--- program CFSteer (robot KUKA KR 30 HA) ---
  BAS (#INITMOV,0)
  BAS (#VEL_PTP,100)
  BAS (#ACC_PTP,20)
  Sollgeschwindigkeit (200.0 mm/s)
  Werkzeug setzen: TOOL 0
  Referenz erstellen.: BASE 0
  $ADVANCE = 5
  $APO.CPTP = 1.000
  $APO.CDIS = 1.000
  Sollgeschwindigkeit (1000.0 mm/s)
  Frame wechseln at (1415.36, -92.38, 659.99) mm, rotated rx -90 ry 0 rz 0 deg
  Werkzeug setzen at (350.64, -42.92, 173.8) mm
  Sollgeschwindigkeit (50.0 mm/s)
  MoveL 2 to (-32.85, -83.54, 62.24) mm, rotated rx 90 ry 17.84 rz 90 deg; joints [-6.49, -82.474, 137.961, 172.14, 55.739, -157.712]
  Sollgeschwindigkeit (50.0 mm/s)
  MoveL 3 to (-32.85, -40.71, 48.45) mm, rotated rx 90 ry 17.84 rz 90 deg; joints [-5.738, -79.848, 139.076, 173.33, 59.399, -158.749]
  MoveL 4 to (-31.86, -40.73, 48.38) mm, rotated rx 90 ry 17.46 rz 90 deg; joints [-5.612, -79.87, 138.999, 173.469, 59.293, -159.191]
  MoveL 5 to (-30.88, -40.75, 48.3) mm, rotated rx 90 ry 17.08 rz 90 deg; joints [-5.486, -79.891, 138.922, 173.609, 59.189, -159.635]
  MoveL 6 to (-29.89, -40.77, 48.23) mm, rotated rx 90 ry 16.7 rz 90 deg; joints [-5.359, -79.911, 138.845, 173.75, 59.085, -160.08]
  MoveL 7 to (-28.9, -40.8, 48.16) mm, rotated rx 90 ry 16.32 rz 90 deg; joints [-5.233, -79.929, 138.768, 173.891, 58.984, -160.524]
  MoveL 8 to (-27.92, -40.82, 48.09) mm, rotated rx 90 ry 15.94 rz 90 deg; joints [-5.106, -79.946, 138.691, 174.033, 58.883, -160.971]
  MoveL 9 to (-26.93, -40.84, 48.02) mm, rotated rx 90 ry 15.56 rz 90 deg; joints [-4.979, -79.961, 138.614, 174.175, 58.784, -161.417]
  MoveL 10 to (-25.95, -40.86, 47.95) mm, rotated rx 90 ry 15.17 rz 90 deg; joints [-4.852, -79.975, 138.537, 174.318, 58.687, -161.866]
  MoveL 11 to (-24.96, -40.88, 47.87) mm, rotated rx 90 ry 14.79 rz 90 deg; joints [-4.725, -79.988, 138.459, 174.461, 58.591, -162.314]
  MoveL 12 to (-23.97, -40.9, 47.8) mm, rotated rx 90 ry 14.41 rz 90 deg; joints [-4.598, -79.999, 138.382, 174.604, 58.496, -162.762]
  MoveL 13 to (-22.99, -40.9, 47.8) mm, rotated rx 90 ry 14.44 rz 90 deg; joints [-4.603, -79.938, 138.311, 174.598, 58.487, -162.729]
  MoveL 14 to (-22, -40.89, 47.81) mm, rotated rx 90 ry 14.47 rz 90 deg; joints [-4.608, -79.877, 138.24, 174.592, 58.478, -162.696]
  MoveL 15 to (-21.01, -40.89, 47.82) mm, rotated rx 90 ry 14.5 rz 90 deg; joints [-4.614, -79.815, 138.17, 174.585, 58.469, -162.663]
  MoveL 16 to (-20.02, -40.89, 47.82) mm, rotated rx 90 ry 14.53 rz 90 deg; joints [-4.618, -79.754, 138.099, 174.579, 58.459, -162.63]
  MoveL 17 to (-19.04, -40.89, 47.83) mm, rotated rx 90 ry 14.56 rz 90 deg; joints [-4.623, -79.693, 138.028, 174.572, 58.45, -162.597]
  MoveL 18 to (-18.05, -40.89, 47.83) mm, rotated rx 90 ry 14.59 rz 90 deg; joints [-4.628, -79.632, 137.957, 174.566, 58.44, -162.564]
  MoveL 19 to (-17.06, -40.89, 47.84) mm, rotated rx 90 ry 14.62 rz 90 deg; joints [-4.633, -79.571, 137.886, 174.56, 58.43, -162.53]
  MoveL 20 to (-16.07, -40.88, 47.84) mm, rotated rx 90 ry 14.64 rz 90 deg; joints [-4.638, -79.51, 137.815, 174.553, 58.421, -162.497]
  MoveL 21 to (-15.09, -40.88, 47.85) mm, rotated rx 90 ry 14.67 rz 90 deg; joints [-4.643, -79.449, 137.744, 174.547, 58.411, -162.464]
  MoveL 22 to (-14.11, -40.84, 47.99) mm, rotated rx 90 ry 15.42 rz 90 deg; joints [-4.875, -79.262, 137.685, 174.282, 58.551, -161.593]
  MoveL 23 to (-13.13, -40.8, 48.13) mm, rotated rx 90 ry 16.16 rz 90 deg; joints [-5.105, -79.07, 137.626, 174.022, 58.695, -160.725]
  MoveL 24 to (-12.15, -40.76, 48.27) mm, rotated rx 90 ry 16.9 rz 90 deg; joints [-5.334, -78.873, 137.566, 173.764, 58.843, -159.86]
  MoveL 25 to (-11.18, -40.72, 48.41) mm, rotated rx 90 ry 17.65 rz 90 deg; joints [-5.56, -78.673, 137.506, 173.509, 58.996, -158.998]
  MoveL 26 to (-10.2, -40.67, 48.55) mm, rotated rx 90 ry 18.39 rz 90 deg; joints [-5.785, -78.468, 137.446, 173.258, 59.153, -158.14]
  MoveL 27 to (-9.22, -40.63, 48.69) mm, rotated rx 90 ry 19.14 rz 90 deg; joints [-6.007, -78.259, 137.385, 173.01, 59.314, -157.285]
  MoveL 28 to (-8.24, -40.58, 48.83) mm, rotated rx 90 ry 19.88 rz 90 deg; joints [-6.228, -78.045, 137.323, 172.766, 59.479, -156.432]
  MoveL 29 to (-7.26, -40.53, 48.96) mm, rotated rx 90 ry 20.62 rz 90 deg; joints [-6.446, -77.828, 137.262, 172.525, 59.647, -155.585]
  MoveL 30 to (-6.28, -40.48, 49.1) mm, rotated rx 90 ry 21.37 rz 90 deg; joints [-6.662, -77.607, 137.2, 172.287, 59.82, -154.739]
  MoveL 31 to (-5.38, -40.38, 49.34) mm, rotated rx 90 ry 22.67 rz 90 deg; joints [-7.042, -77.252, 137.149, 171.874, 60.146, -153.264]
  MoveL 32 to (-4.47, -40.28, 49.57) mm, rotated rx 90 ry 23.98 rz 90 deg; joints [-7.415, -76.885, 137.096, 171.471, 60.485, -151.8]
  MoveL 33 to (-3.56, -40.17, 49.8) mm, rotated rx 90 ry 25.28 rz 90 deg; joints [-7.782, -76.505, 137.042, 171.079, 60.835, -150.347]
  MoveL 34 to (-2.66, -40.06, 50.03) mm, rotated rx 90 ry 26.58 rz 90 deg; joints [-8.143, -76.113, 136.987, 170.698, 61.196, -148.903]
  MoveL 35 to (-1.75, -39.94, 50.26) mm, rotated rx 90 ry 27.89 rz 90 deg; joints [-8.497, -75.708, 136.93, 170.327, 61.567, -147.472]
  MoveL 36 to (-0.84, -39.82, 50.49) mm, rotated rx 90 ry 29.19 rz 90 deg; joints [-8.844, -75.292, 136.872, 169.968, 61.948, -146.052]
  MoveL 37 to (0.05, -39.66, 50.77) mm, rotated rx 90 ry 30.83 rz 90 deg; joints [-9.272, -74.765, 136.814, 169.529, 62.446, -144.283]
  MoveL 38 to (0.93, -39.49, 51.04) mm, rotated rx 90 ry 32.47 rz 90 deg; joints [-9.689, -74.22, 136.754, 169.108, 62.958, -142.53]
  MoveL 39 to (1.82, -39.31, 51.31) mm, rotated rx 90 ry 34.11 rz 90 deg; joints [-10.094, -73.657, 136.691, 168.704, 63.484, -140.795]
  MoveL 40 to (2.71, -39.13, 51.57) mm, rotated rx 90 ry 35.75 rz 90 deg; joints [-10.488, -73.076, 136.624, 168.317, 64.023, -139.077]
  MoveL 41 to (3.6, -38.94, 51.83) mm, rotated rx 90 ry 37.39 rz 90 deg; joints [-10.87, -72.479, 136.554, 167.948, 64.574, -137.376]
  MoveL 42 to (4.49, -38.74, 52.08) mm, rotated rx 90 ry 39.02 rz 90 deg; joints [-11.239, -71.866, 136.481, 167.595, 65.136, -135.691]
  MoveL 43 to (5.36, -38.51, 52.36) mm, rotated rx 90 ry 40.85 rz 90 deg; joints [-11.636, -71.171, 136.404, 167.222, 65.775, -133.838]
  MoveL 44 to (6.24, -38.27, 52.62) mm, rotated rx 90 ry 42.67 rz 90 deg; joints [-12.018, -70.457, 136.322, 166.869, 66.426, -132.003]
  MoveL 45 to (7.12, -38.03, 52.88) mm, rotated rx 90 ry 44.49 rz 90 deg; joints [-12.383, -69.726, 136.235, 166.537, 67.088, -130.188]
  MoveL 46 to (7.99, -37.77, 53.13) mm, rotated rx 90 ry 46.31 rz 90 deg; joints [-12.733, -68.977, 136.144, 166.224, 67.759, -128.39]
  MoveL 47 to (8.87, -37.51, 53.38) mm, rotated rx 90 ry 48.13 rz 90 deg; joints [-13.066, -68.212, 136.047, 165.932, 68.438, -126.609]
  MoveL 48 to (9.75, -37.24, 53.61) mm, rotated rx 90 ry 49.95 rz 90 deg; joints [-13.383, -67.431, 135.945, 165.658, 69.125, -124.844]
  MoveL 49 to (10.62, -36.95, 53.85) mm, rotated rx 90 ry 51.84 rz 90 deg; joints [-13.694, -66.608, 135.837, 165.394, 69.846, -123.031]
  MoveL 50 to (11.5, -36.66, 54.07) mm, rotated rx 90 ry 53.73 rz 90 deg; joints [-13.987, -65.769, 135.723, 165.15, 70.572, -121.233]
  MoveL 51 to (12.37, -36.35, 54.28) mm, rotated rx 90 ry 55.62 rz 90 deg; joints [-14.261, -64.917, 135.603, 164.926, 71.303, -119.45]
  MoveL 52 to (13.24, -36.04, 54.49) mm, rotated rx 90 ry 57.5 rz 90 deg; joints [-14.518, -64.051, 135.476, 164.721, 72.039, -117.681]
  MoveL 53 to (14.12, -35.73, 54.68) mm, rotated rx 90 ry 59.39 rz 90 deg; joints [-14.755, -63.175, 135.344, 164.535, 72.776, -115.925]
  MoveL 54 to (14.99, -35.41, 54.87) mm, rotated rx 90 ry 61.28 rz 90 deg; joints [-14.974, -62.286, 135.206, 164.368, 73.517, -114.18]
  MoveL 55 to (15.87, -35.1, 55.03) mm, rotated rx 90 ry 63.05 rz 90 deg; joints [-15.161, -61.443, 135.067, 164.229, 74.209, -112.554]
  MoveL 56 to (16.74, -34.79, 55.18) mm, rotated rx 90 ry 64.82 rz 90 deg; joints [-15.332, -60.592, 134.922, 164.105, 74.901, -110.937]
  MoveL 57 to (17.61, -34.47, 55.32) mm, rotated rx 90 ry 66.59 rz 90 deg; joints [-15.486, -59.734, 134.772, 163.998, 75.593, -109.327]
  MoveL 58 to (18.49, -34.15, 55.46) mm, rotated rx 90 ry 68.36 rz 90 deg; joints [-15.624, -58.87, 134.616, 163.905, 76.283, -107.725]
  MoveL 59 to (19.36, -33.82, 55.58) mm, rotated rx 90 ry 70.13 rz 90 deg; joints [-15.744, -58.001, 134.456, 163.829, 76.972, -106.129]
  MoveL 60 to (20.23, -33.49, 55.69) mm, rotated rx 90 ry 71.9 rz 90 deg; joints [-15.848, -57.128, 134.289, 163.767, 77.657, -104.538]
  MoveL 61 to (21.12, -33.23, 55.78) mm, rotated rx 90 ry 73.31 rz 90 deg; joints [-15.916, -56.424, 134.139, 163.73, 78.193, -103.273]
  MoveL 62 to (22, -32.97, 55.85) mm, rotated rx 90 ry 74.72 rz 90 deg; joints [-15.973, -55.719, 133.986, 163.704, 78.726, -102.01]
  MoveL 63 to (22.88, -32.7, 55.92) mm, rotated rx 90 ry 76.13 rz 90 deg; joints [-16.02, -55.013, 133.83, 163.686, 79.256, -100.749]
  MoveL 64 to (23.77, -32.43, 55.98) mm, rotated rx 90 ry 77.54 rz 90 deg; joints [-16.056, -54.307, 133.67, 163.678, 79.783, -99.49]
  MoveL 65 to (24.65, -32.16, 56.04) mm, rotated rx 90 ry 78.95 rz 90 deg; joints [-16.082, -53.6, 133.508, 163.679, 80.307, -98.231]
  MoveL 66 to (25.53, -31.89, 56.09) mm, rotated rx 90 ry 80.36 rz 90 deg; joints [-16.096, -52.893, 133.342, 163.689, 80.827, -96.974]
  MoveL 67 to (26.46, -31.75, 56.11) mm, rotated rx 90 ry 81.07 rz 90 deg; joints [-16.093, -52.524, 133.222, 163.704, 81.065, -96.333]
  MoveL 68 to (27.39, -31.61, 56.13) mm, rotated rx 90 ry 81.78 rz 90 deg; joints [-16.087, -52.155, 133.1, 163.721, 81.303, -95.692]
  MoveL 69 to (28.32, -31.47, 56.15) mm, rotated rx 90 ry 82.49 rz 90 deg; joints [-16.078, -51.786, 132.978, 163.74, 81.539, -95.051]
  MoveL 70 to (29.25, -31.33, 56.17) mm, rotated rx 90 ry 83.2 rz 90 deg; joints [-16.067, -51.418, 132.856, 163.762, 81.774, -94.409]
  MoveL 71 to (30.18, -31.19, 56.19) mm, rotated rx 90 ry 83.92 rz 90 deg; joints [-16.053, -51.052, 132.733, 163.785, 82.008, -93.768]
  MoveL 72 to (31.11, -31.05, 56.2) mm, rotated rx 90 ry 84.63 rz 90 deg; joints [-16.036, -50.685, 132.608, 163.812, 82.24, -93.125]
  MoveL 73 to (31.98, -31.11, 56.2) mm, rotated rx 90 ry 84.31 rz 90 deg; joints [-16.026, -50.818, 132.569, 163.815, 82.074, -93.398]
  MoveL 74 to (32.86, -31.18, 56.19) mm, rotated rx 90 ry 83.99 rz 90 deg; joints [-16.016, -50.951, 132.53, 163.819, 81.907, -93.671]
  MoveL 75 to (33.73, -31.24, 56.18) mm, rotated rx 90 ry 83.67 rz 90 deg; joints [-16.005, -51.084, 132.49, 163.823, 81.742, -93.943]
  MoveL 76 to (34.6, -31.3, 56.17) mm, rotated rx 90 ry 83.35 rz 90 deg; joints [-15.993, -51.216, 132.45, 163.828, 81.576, -94.216]
  MoveL 77 to (35.48, -31.36, 56.17) mm, rotated rx 90 ry 83.03 rz 90 deg; joints [-15.981, -51.348, 132.41, 163.833, 81.41, -94.489]
  MoveL 78 to (36.35, -31.43, 56.16) mm, rotated rx 90 ry 82.71 rz 90 deg; joints [-15.968, -51.479, 132.37, 163.838, 81.245, -94.762]
  MoveL 79 to (37.22, -31.49, 56.15) mm, rotated rx 90 ry 82.39 rz 90 deg; joints [-15.955, -51.61, 132.329, 163.844, 81.079, -95.035]
  MoveL 80 to (38.14, -31.69, 56.12) mm, rotated rx 90 ry 81.34 rz 90 deg; joints [-15.935, -52.089, 132.339, 163.843, 80.628, -95.954]
  MoveL 81 to (39.06, -31.9, 56.09) mm, rotated rx 90 ry 80.3 rz 90 deg; joints [-15.909, -52.566, 132.346, 163.847, 80.176, -96.874]
  MoveL 82 to (39.98, -32.1, 56.05) mm, rotated rx 90 ry 79.25 rz 90 deg; joints [-15.878, -53.042, 132.353, 163.856, 79.723, -97.796]
  MoveL 83 to (40.9, -32.3, 56.01) mm, rotated rx 90 ry 78.2 rz 90 deg; joints [-15.84, -53.516, 132.357, 163.87, 79.27, -98.718]
  MoveL 84 to (41.81, -32.5, 55.97) mm, rotated rx 90 ry 77.15 rz 90 deg; joints [-15.797, -53.988, 132.359, 163.889, 78.816, -99.641]
  MoveL 85 to (42.73, -32.7, 55.92) mm, rotated rx 90 ry 76.1 rz 90 deg; joints [-15.748, -54.458, 132.36, 163.912, 78.362, -100.566]
  MoveL 86 to (43.65, -32.9, 55.87) mm, rotated rx 90 ry 75.06 rz 90 deg; joints [-15.694, -54.926, 132.358, 163.941, 77.908, -101.493]
  MoveL 87 to (44.61, -32.99, 55.84) mm, rotated rx 90 ry 74.56 rz 90 deg; joints [-15.659, -55.131, 132.318, 163.962, 77.67, -101.928]
  MoveL 88 to (45.57, -33.09, 55.82) mm, rotated rx 90 ry 74.06 rz 90 deg; joints [-15.623, -55.336, 132.277, 163.984, 77.432, -102.364]
  MoveL 89 to (46.52, -33.18, 55.79) mm, rotated rx 90 ry 73.56 rz 90 deg; joints [-15.585, -55.54, 132.236, 164.007, 77.194, -102.8]
  MoveL 90 to (47.48, -33.28, 55.76) mm, rotated rx 90 ry 73.07 rz 90 deg; joints [-15.547, -55.742, 132.194, 164.031, 76.956, -103.236]
  MoveL 91 to (48.44, -33.37, 55.73) mm, rotated rx 90 ry 72.57 rz 90 deg; joints [-15.507, -55.944, 132.152, 164.056, 76.719, -103.673]
  MoveL 92 to (49.4, -33.46, 55.7) mm, rotated rx 90 ry 72.08 rz 90 deg; joints [-15.466, -56.145, 132.109, 164.082, 76.482, -104.111]
  MoveL 93 to (50.35, -33.55, 55.67) mm, rotated rx 90 ry 71.58 rz 90 deg; joints [-15.424, -56.345, 132.066, 164.109, 76.245, -104.55]
  MoveL 94 to (51.31, -33.44, 55.71) mm, rotated rx 90 ry 72.18 rz 90 deg; joints [-15.447, -56.037, 131.96, 164.099, 76.442, -103.999]
  MoveL 95 to (52.26, -33.33, 55.75) mm, rotated rx 90 ry 72.78 rz 90 deg; joints [-15.468, -55.728, 131.853, 164.09, 76.638, -103.448]
  MoveL 96 to (53.21, -33.22, 55.78) mm, rotated rx 90 ry 73.39 rz 90 deg; joints [-15.488, -55.419, 131.746, 164.083, 76.832, -102.898]
  MoveL 97 to (54.16, -33.1, 55.81) mm, rotated rx 90 ry 73.99 rz 90 deg; joints [-15.505, -55.11, 131.638, 164.078, 77.027, -102.348]
  MoveL 98 to (55.12, -32.99, 55.85) mm, rotated rx 90 ry 74.59 rz 90 deg; joints [-15.521, -54.802, 131.53, 164.074, 77.221, -101.798]
  MoveL 99 to (56.07, -32.88, 55.88) mm, rotated rx 90 ry 75.19 rz 90 deg; joints [-15.535, -54.493, 131.421, 164.073, 77.414, -101.249]
  MoveL 100 to (57.02, -32.76, 55.91) mm, rotated rx 90 ry 75.8 rz 90 deg; joints [-15.547, -54.185, 131.312, 164.073, 77.605, -100.7]
  MoveL 101 to (57.94, -32.56, 55.95) mm, rotated rx 90 ry 76.82 rz 90 deg; joints [-15.572, -53.681, 131.177, 164.069, 77.962, -99.772]
  MoveL 102 to (58.86, -32.37, 56) mm, rotated rx 90 ry 77.85 rz 90 deg; joints [-15.591, -53.177, 131.04, 164.07, 78.317, -98.846]
  MoveL 103 to (59.77, -32.17, 56.04) mm, rotated rx 90 ry 78.87 rz 90 deg; joints [-15.605, -52.672, 130.902, 164.076, 78.67, -97.92]
  MoveL 104 to (60.69, -31.97, 56.08) mm, rotated rx 90 ry 79.9 rz 90 deg; joints [-15.614, -52.169, 130.763, 164.087, 79.02, -96.995]
  MoveL 105 to (61.61, -31.77, 56.11) mm, rotated rx 90 ry 80.92 rz 90 deg; joints [-15.617, -51.665, 130.622, 164.103, 79.369, -96.069]
  MoveL 106 to (62.52, -31.58, 56.14) mm, rotated rx 90 ry 81.95 rz 90 deg; joints [-15.614, -51.163, 130.48, 164.124, 79.715, -95.145]
  MoveL 107 to (63.44, -31.38, 56.17) mm, rotated rx 90 ry 82.97 rz 90 deg; joints [-15.607, -50.661, 130.336, 164.149, 80.06, -94.22]
  MoveL 108 to (64.31, -31.34, 56.17) mm, rotated rx 90 ry 83.18 rz 90 deg; joints [-15.596, -50.54, 130.255, 164.162, 80.098, -94.022]
  MoveL 109 to (65.17, -31.29, 56.17) mm, rotated rx 90 ry 83.4 rz 90 deg; joints [-15.584, -50.42, 130.175, 164.176, 80.136, -93.825]
  MoveL 110 to (66.03, -31.25, 56.18) mm, rotated rx 90 ry 83.61 rz 90 deg; joints [-15.573, -50.299, 130.094, 164.19, 80.174, -93.627]
  MoveL 111 to (66.9, -31.21, 56.19) mm, rotated rx 90 ry 83.82 rz 90 deg; joints [-15.561, -50.179, 130.014, 164.203, 80.211, -93.429]
  MoveL 112 to (67.76, -31.17, 56.19) mm, rotated rx 90 ry 84.03 rz 90 deg; joints [-15.549, -50.058, 129.933, 164.217, 80.249, -93.231]
  MoveL 113 to (68.63, -31.13, 56.19) mm, rotated rx 90 ry 84.24 rz 90 deg; joints [-15.537, -49.938, 129.853, 164.232, 80.286, -93.033]
  MoveL 114 to (69.49, -31.09, 56.2) mm, rotated rx 90 ry 84.45 rz 90 deg; joints [-15.524, -49.819, 129.772, 164.246, 80.323, -92.835]
  MoveL 115 to (70.41, -31.25, 56.18) mm, rotated rx 90 ry 83.65 rz 90 deg; joints [-15.516, -50.166, 129.763, 164.238, 79.98, -93.541]
  MoveL 116 to (71.33, -31.4, 56.16) mm, rotated rx 90 ry 82.84 rz 90 deg; joints [-15.504, -50.513, 129.753, 164.232, 79.637, -94.248]
  MoveL 117 to (72.26, -31.56, 56.14) mm, rotated rx 90 ry 82.04 rz 90 deg; joints [-15.489, -50.859, 129.743, 164.23, 79.292, -94.955]
  MoveL 118 to (73.18, -31.71, 56.12) mm, rotated rx 90 ry 81.24 rz 90 deg; joints [-15.47, -51.204, 129.731, 164.23, 78.948, -95.664]
  MoveL 119 to (74.1, -31.87, 56.09) mm, rotated rx 90 ry 80.43 rz 90 deg; joints [-15.448, -51.549, 129.718, 164.233, 78.603, -96.373]
  MoveL 120 to (75.03, -32.02, 56.07) mm, rotated rx 90 ry 79.63 rz 90 deg; joints [-15.423, -51.892, 129.704, 164.239, 78.258, -97.082]
  MoveL 121 to (75.91, -32.31, 56.01) mm, rotated rx 90 ry 78.17 rz 90 deg; joints [-15.379, -52.536, 129.737, 164.248, 77.667, -98.381]
  MoveL 122 to (76.79, -32.59, 55.95) mm, rotated rx 90 ry 76.71 rz 90 deg; joints [-15.325, -53.177, 129.765, 164.267, 77.074, -99.683]
  MoveL 123 to (77.67, -32.86, 55.88) mm, rotated rx 90 ry 75.25 rz 90 deg; joints [-15.259, -53.814, 129.791, 164.295, 76.48, -100.988]
  MoveL 124 to (78.55, -33.14, 55.8) mm, rotated rx 90 ry 73.79 rz 90 deg; joints [-15.183, -54.449, 129.813, 164.333, 75.886, -102.297]
  MoveL 125 to (79.43, -33.41, 55.72) mm, rotated rx 90 ry 72.33 rz 90 deg; joints [-15.095, -55.079, 129.831, 164.38, 75.291, -103.61]
  MoveL 126 to (80.31, -33.69, 55.63) mm, rotated rx 90 ry 70.87 rz 90 deg; joints [-14.997, -55.704, 129.846, 164.438, 74.696, -104.926]
  MoveL 127 to (81.19, -34.02, 55.51) mm, rotated rx 90 ry 69.08 rz 90 deg; joints [-14.865, -56.471, 129.876, 164.519, 73.975, -106.551]
  MoveL 128 to (82.06, -34.34, 55.38) mm, rotated rx 90 ry 67.28 rz 90 deg; joints [-14.717, -57.231, 129.9, 164.616, 73.255, -108.183]
  MoveL 129 to (82.93, -34.67, 55.24) mm, rotated rx 90 ry 65.49 rz 90 deg; joints [-14.553, -57.982, 129.919, 164.727, 72.536, -109.824]
  MoveL 130 to (83.81, -34.98, 55.09) mm, rotated rx 90 ry 63.7 rz 90 deg; joints [-14.373, -58.723, 129.933, 164.855, 71.819, -111.475]
  MoveL 131 to (84.68, -35.3, 54.92) mm, rotated rx 90 ry 61.91 rz 90 deg; joints [-14.177, -59.453, 129.941, 164.997, 71.105, -113.135]
  MoveL 132 to (85.55, -35.61, 54.75) mm, rotated rx 90 ry 60.11 rz 90 deg; joints [-13.966, -60.173, 129.945, 165.156, 70.394, -114.807]
  MoveL 133 to (86.51, -35.95, 54.55) mm, rotated rx 90 ry 58.07 rz 90 deg; joints [-13.706, -60.981, 129.945, 165.356, 69.59, -116.727]
  MoveL 134 to (87.46, -36.29, 54.33) mm, rotated rx 90 ry 56.02 rz 90 deg; joints [-13.427, -61.772, 129.939, 165.577, 68.793, -118.664]
  MoveL 135 to (88.42, -36.62, 54.1) mm, rotated rx 90 ry 53.98 rz 90 deg; joints [-13.129, -62.546, 129.926, 165.82, 68.003, -120.618]
  MoveL 136 to (89.37, -36.94, 53.86) mm, rotated rx 90 ry 51.93 rz 90 deg; joints [-12.811, -63.301, 129.907, 166.085, 67.222, -122.59]
  MoveL 137 to (90.32, -37.25, 53.6) mm, rotated rx 90 ry 49.89 rz 90 deg; joints [-12.474, -64.036, 129.882, 166.372, 66.451, -124.581]
  MoveL 138 to (91.28, -37.55, 53.34) mm, rotated rx 90 ry 47.84 rz 90 deg; joints [-12.119, -64.751, 129.851, 166.682, 65.691, -126.593]
  MoveL 139 to (92.23, -37.84, 53.06) mm, rotated rx 90 ry 45.8 rz 90 deg; joints [-11.745, -65.445, 129.814, 167.014, 64.943, -128.626]
  MoveL 140 to (93.19, -38.13, 52.78) mm, rotated rx 90 ry 43.75 rz 90 deg; joints [-11.354, -66.116, 129.771, 167.37, 64.209, -130.681]
  MoveL 141 to (94.15, -38.37, 52.52) mm, rotated rx 90 ry 41.92 rz 90 deg; joints [-10.987, -66.693, 129.719, 167.711, 63.559, -132.544]
  MoveL 142 to (95.12, -38.61, 52.24) mm, rotated rx 90 ry 40.08 rz 90 deg; joints [-10.606, -67.25, 129.663, 168.07, 62.923, -134.426]
  MoveL 143 to (96.08, -38.84, 51.96) mm, rotated rx 90 ry 38.25 rz 90 deg; joints [-10.212, -67.788, 129.603, 168.449, 62.3, -136.327]
  MoveL 144 to (97.05, -39.05, 51.68) mm, rotated rx 90 ry 36.41 rz 90 deg; joints [-9.805, -68.305, 129.539, 168.847, 61.693, -138.248]
  MoveL 145 to (98.01, -39.26, 51.38) mm, rotated rx 90 ry 34.58 rz 90 deg; joints [-9.386, -68.8, 129.471, 169.264, 61.102, -140.188]
  MoveL 146 to (98.98, -39.46, 51.09) mm, rotated rx 90 ry 32.74 rz 90 deg; joints [-8.955, -69.274, 129.4, 169.7, 60.527, -142.149]
  MoveL 147 to (99.94, -39.65, 50.78) mm, rotated rx 90 ry 30.91 rz 90 deg; joints [-8.512, -69.725, 129.326, 170.156, 59.97, -144.13]
  MoveL 148 to (100.91, -39.83, 50.47) mm, rotated rx 90 ry 29.07 rz 90 deg; joints [-8.057, -70.154, 129.248, 170.631, 59.431, -146.132]
  MoveL 149 to (101.91, -39.95, 50.24) mm, rotated rx 90 ry 27.77 rz 90 deg; joints [-7.727, -70.429, 129.167, 170.981, 59.053, -147.563]
  MoveL 150 to (102.9, -40.07, 50.01) mm, rotated rx 90 ry 26.47 rz 90 deg; joints [-7.391, -70.691, 129.085, 171.34, 58.686, -149.004]
  MoveL 151 to (103.9, -40.18, 49.78) mm, rotated rx 90 ry 25.17 rz 90 deg; joints [-7.05, -70.942, 129.001, 171.709, 58.329, -150.457]
  MoveL 152 to (104.89, -40.29, 49.55) mm, rotated rx 90 ry 23.87 rz 90 deg; joints [-6.704, -71.18, 128.916, 172.086, 57.983, -151.918]
  MoveL 153 to (105.89, -40.39, 49.32) mm, rotated rx 90 ry 22.57 rz 90 deg; joints [-6.354, -71.406, 128.829, 172.472, 57.649, -153.389]
  MoveL 154 to (106.89, -40.48, 49.08) mm, rotated rx 90 ry 21.26 rz 90 deg; joints [-6, -71.619, 128.742, 172.866, 57.326, -154.87]
  MoveL 155 to (107.88, -40.57, 48.84) mm, rotated rx 90 ry 19.96 rz 90 deg; joints [-5.642, -71.82, 128.653, 173.269, 57.015, -156.36]
  MoveL 156 to (108.88, -40.66, 48.6) mm, rotated rx 90 ry 18.66 rz 90 deg; joints [-5.28, -72.008, 128.564, 173.68, 56.716, -157.859]
  MoveL 157 to (109.79, -40.69, 48.51) mm, rotated rx 90 ry 18.16 rz 90 deg; joints [-5.135, -72.05, 128.488, 173.845, 56.591, -158.446]
  MoveL 158 to (110.7, -40.72, 48.41) mm, rotated rx 90 ry 17.65 rz 90 deg; joints [-4.99, -72.091, 128.413, 174.01, 56.467, -159.035]
  MoveL 159 to (111.61, -40.75, 48.32) mm, rotated rx 90 ry 17.14 rz 90 deg; joints [-4.845, -72.129, 128.337, 174.176, 56.345, -159.624]
  MoveL 160 to (112.52, -40.78, 48.22) mm, rotated rx 90 ry 16.63 rz 90 deg; joints [-4.699, -72.165, 128.262, 174.344, 56.226, -160.215]
  MoveL 161 to (113.43, -40.81, 48.12) mm, rotated rx 90 ry 16.13 rz 90 deg; joints [-4.553, -72.199, 128.186, 174.512, 56.108, -160.806]
  MoveL 162 to (114.34, -40.84, 48.03) mm, rotated rx 90 ry 15.62 rz 90 deg; joints [-4.407, -72.232, 128.11, 174.682, 55.992, -161.401]
  MoveL 163 to (115.25, -40.86, 47.93) mm, rotated rx 90 ry 15.11 rz 90 deg; joints [-4.26, -72.262, 128.033, 174.852, 55.879, -161.995]
  MoveL 164 to (116.16, -40.89, 47.84) mm, rotated rx 90 ry 14.61 rz 90 deg; joints [-4.113, -72.29, 127.957, 175.024, 55.768, -162.591]
  MoveL 165 to (117.07, -40.91, 47.74) mm, rotated rx 90 ry 14.1 rz 90 deg; joints [-3.965, -72.316, 127.88, 175.196, 55.658, -163.187]
  MoveL 166 to (117.99, -40.91, 47.76) mm, rotated rx 90 ry 14.17 rz 90 deg; joints [-3.984, -72.256, 127.811, 175.172, 55.65, -163.097]
  MoveL 167 to (118.9, -40.9, 47.77) mm, rotated rx 90 ry 14.25 rz 90 deg; joints [-4.003, -72.197, 127.742, 175.149, 55.641, -163.006]
  MoveL 168 to (119.81, -40.9, 47.78) mm, rotated rx 90 ry 14.33 rz 90 deg; joints [-4.022, -72.137, 127.673, 175.126, 55.633, -162.915]
  MoveL 169 to (120.73, -40.9, 47.8) mm, rotated rx 90 ry 14.41 rz 90 deg; joints [-4.041, -72.077, 127.603, 175.102, 55.624, -162.824]
  MoveL 170 to (121.64, -40.89, 47.81) mm, rotated rx 90 ry 14.48 rz 90 deg; joints [-4.059, -72.017, 127.534, 175.079, 55.616, -162.733]
  MoveL 171 to (122.55, -40.89, 47.83) mm, rotated rx 90 ry 14.56 rz 90 deg; joints [-4.078, -71.957, 127.464, 175.056, 55.607, -162.643]
  MoveL 172 to (123.47, -40.88, 47.84) mm, rotated rx 90 ry 14.64 rz 90 deg; joints [-4.097, -71.897, 127.395, 175.033, 55.598, -162.552]
  MoveL 173 to (124.38, -40.88, 47.86) mm, rotated rx 90 ry 14.71 rz 90 deg; joints [-4.116, -71.837, 127.326, 175.009, 55.59, -162.46]
  MoveL 174 to (125.3, -40.88, 47.87) mm, rotated rx 90 ry 14.79 rz 90 deg; joints [-4.134, -71.777, 127.256, 174.986, 55.581, -162.369]
  MoveL 175 to (126.21, -40.86, 47.94) mm, rotated rx 90 ry 15.16 rz 90 deg; joints [-4.235, -71.673, 127.19, 174.867, 55.624, -161.934]
  MoveL 176 to (127.12, -40.84, 48.01) mm, rotated rx 90 ry 15.53 rz 90 deg; joints [-4.336, -71.568, 127.124, 174.747, 55.668, -161.499]
  MoveL 177 to (128.03, -40.82, 48.08) mm, rotated rx 90 ry 15.9 rz 90 deg; joints [-4.436, -71.462, 127.058, 174.629, 55.713, -161.064]
  MoveL 178 to (128.94, -40.8, 48.15) mm, rotated rx 90 ry 16.27 rz 90 deg; joints [-4.536, -71.356, 126.992, 174.511, 55.759, -160.63]
  MoveL 179 to (129.86, -40.78, 48.22) mm, rotated rx 90 ry 16.64 rz 90 deg; joints [-4.635, -71.248, 126.926, 174.394, 55.805, -160.197]
  MoveL 180 to (130.77, -40.76, 48.29) mm, rotated rx 90 ry 17.02 rz 90 deg; joints [-4.734, -71.14, 126.859, 174.277, 55.852, -159.764]
  MoveL 181 to (131.68, -40.74, 48.36) mm, rotated rx 90 ry 17.39 rz 90 deg; joints [-4.832, -71.031, 126.793, 174.161, 55.9, -159.332]
  MoveL 182 to (132.59, -40.71, 48.43) mm, rotated rx 90 ry 17.76 rz 90 deg; joints [-4.93, -70.921, 126.726, 174.046, 55.949, -158.9]
  MoveL 183 to (133.51, -40.69, 48.5) mm, rotated rx 90 ry 18.13 rz 90 deg; joints [-5.027, -70.81, 126.659, 173.932, 55.999, -158.469]
  MoveL 184 to (134.42, -40.67, 48.56) mm, rotated rx 90 ry 18.43 rz 90 deg; joints [-5.106, -70.71, 126.591, 173.84, 56.035, -158.119]
  MoveL 185 to (135.33, -40.65, 48.61) mm, rotated rx 90 ry 18.73 rz 90 deg; joints [-5.184, -70.609, 126.524, 173.749, 56.073, -157.767]
  MoveL 186 to (136.25, -40.63, 48.67) mm, rotated rx 90 ry 19.04 rz 90 deg; joints [-5.262, -70.508, 126.456, 173.657, 56.11, -157.416]
  MoveL 187 to (137.16, -40.62, 48.73) mm, rotated rx 90 ry 19.34 rz 90 deg; joints [-5.339, -70.407, 126.388, 173.567, 56.149, -157.066]
  MoveL 188 to (138.07, -40.59, 48.78) mm, rotated rx 90 ry 19.64 rz 90 deg; joints [-5.416, -70.305, 126.32, 173.477, 56.187, -156.716]
  MoveL 189 to (138.98, -40.58, 48.84) mm, rotated rx 90 ry 19.95 rz 90 deg; joints [-5.493, -70.202, 126.252, 173.387, 56.226, -156.366]
  MoveL 190 to (139.9, -40.55, 48.89) mm, rotated rx 90 ry 20.25 rz 90 deg; joints [-5.57, -70.099, 126.183, 173.298, 56.266, -156.017]
  MoveL 191 to (140.81, -40.53, 48.95) mm, rotated rx 90 ry 20.55 rz 90 deg; joints [-5.646, -69.996, 126.115, 173.21, 56.306, -155.669]
  MoveL 192 to (141.72, -40.51, 49.01) mm, rotated rx 90 ry 20.85 rz 90 deg; joints [-5.721, -69.892, 126.047, 173.122, 56.346, -155.322]
  MoveL 193 to (142.4, -40.79, 48.17) mm, rotated rx 90 ry 16.38 rz 90 deg; joints [-4.515, -70.63, 125.949, 174.515, 55.442, -160.499]
  MoveL 194 to (143.07, -41.01, 47.32) mm, rotated rx 90 ry 11.91 rz 90 deg; joints [-3.266, -71.227, 125.841, 175.996, 54.68, -165.771]
  MoveL 195 to (143.75, -41.16, 46.46) mm, rotated rx 90 ry 7.44 rz 90 deg; joints [-1.981, -71.678, 125.723, 177.553, 54.07, -171.124]
  MoveL 196 to (144.43, -41.23, 45.58) mm, rotated rx 90 ry 2.97 rz 90 deg; joints [-0.67, -71.982, 125.598, 179.168, 53.619, -176.537]
  MoveL 197 to (145.1, -41.25, 44.7) mm, rotated rx 90 ry 0 rz 90 deg; joints [0.224, -72.088, 125.494, -179.721, 53.406, 179.834]
  MoveL 198 to (141.7, -41.25, 42.87) mm, rotated rx 90 ry 0 rz 90 deg; joints [0.311, -72.273, 125.758, -179.612, 53.486, 179.769]
  MoveL 199 to (137.91, -41.25, 41.96) mm, rotated rx 90 ry 0 rz 90 deg; joints [0.355, -72.478, 126.051, -179.558, 53.573, 179.738]
  MoveL 200 to (134, -41.25, 41.48) mm, rotated rx 90 ry 0 rz 90 deg; joints [0.379, -72.691, 126.353, -179.529, 53.663, 179.721]
  MoveL 201 to (130.09, -41.25, 41.08) mm, rotated rx 90 ry 0 rz 90 deg; joints [0.4, -72.903, 126.655, -179.505, 53.752, 179.707]
  MoveL 202 to (126.21, -41.25, 40.71) mm, rotated rx 90 ry 0 rz 90 deg; joints [0.419, -73.115, 126.954, -179.481, 53.84, 179.694]
  MoveL 203 to (118.64, -41.25, 39.88) mm, rotated rx 90 ry 0 rz 90 deg; joints [0.461, -73.528, 127.535, -179.43, 54.008, 179.665]
  MoveL 204 to (111.13, -41.25, 38.67) mm, rotated rx 90 ry 0 rz 90 deg; joints [0.523, -73.939, 128.109, -179.355, 54.172, 179.623]
  MoveL 205 to (104.5, -41.25, 37.04) mm, rotated rx 90 ry 0 rz 90 deg; joints [0.605, -74.302, 128.613, -179.255, 54.314, 179.565]
  MoveL 206 to (98.04, -41.25, 34.74) mm, rotated rx 90 ry 0 rz 90 deg; joints [0.721, -74.656, 129.102, -179.113, 54.45, 179.485]
  MoveL 207 to (91.88, -41.25, 31.62) mm, rotated rx 90 ry 0 rz 90 deg; joints [0.879, -74.993, 129.566, -178.922, 54.578, 179.375]
  MoveL 208 to (86.28, -41.25, 27.66) mm, rotated rx 90 ry 0 rz 90 deg; joints [1.079, -75.299, 129.984, -178.678, 54.692, 179.236]
  MoveL 209 to (80.96, -41.25, 22.17) mm, rotated rx 90 ry 0 rz 90 deg; joints [1.356, -75.587, 130.376, -178.34, 54.801, 179.043]
  MoveL 210 to (76.3, -41.25, 15.86) mm, rotated rx 90 ry 0 rz 90 deg; joints [1.677, -75.837, 130.714, -177.95, 54.895, 178.821]
  MoveL 211 to (75.7, -41.25, 15.02) mm, rotated rx 90 ry 0 rz 90 deg; joints [1.72, -75.868, 130.757, -177.898, 54.907, 178.791]
  MoveL 212 to (75.11, -41.22, 14.18) mm, rotated rx 90 ry -4.2 rz 90 deg; joints [3.049, -75.959, 130.67, -176.267, 54.768, 173.646]
  MoveL 213 to (74.51, -41.13, 13.34) mm, rotated rx 90 ry -8.49 rz 90 deg; joints [4.409, -75.905, 130.577, -174.602, 54.792, 168.391]
  MoveL 214 to (73.92, -40.97, 12.51) mm, rotated rx 90 ry -12.78 rz 90 deg; joints [5.762, -75.702, 130.481, -172.958, 54.983, 163.164]
  MoveL 215 to (73.33, -40.76, 11.71) mm, rotated rx 90 ry -17.03 rz 90 deg; joints [7.085, -75.358, 130.384, -171.375, 55.332, 158.042]
  MoveL 216 to (72.75, -40.48, 10.92) mm, rotated rx 90 ry -21.27 rz 90 deg; joints [8.385, -74.874, 130.285, -169.849, 55.833, 152.988]
  MoveL 217 to (72.17, -40.15, 10.15) mm, rotated rx 90 ry -25.52 rz 90 deg; joints [9.653, -74.253, 130.184, -168.397, 56.477, 148.015]
  MoveL 218 to (71.58, -39.77, 9.42) mm, rotated rx 90 ry -29.76 rz 90 deg; joints [10.881, -73.501, 130.08, -167.03, 57.256, 143.14]
  MoveL 219 to (71.04, -39.35, 8.74) mm, rotated rx 90 ry -33.79 rz 90 deg; joints [12.006, -72.668, 129.976, -165.819, 58.109, 138.604]
  MoveL 220 to (70.5, -38.89, 8.1) mm, rotated rx 90 ry -37.83 rz 90 deg; joints [13.083, -71.724, 129.868, -164.698, 59.064, 134.168]
  MoveL 221 to (69.96, -38.38, 7.49) mm, rotated rx 90 ry -41.86 rz 90 deg; joints [14.108, -70.676, 129.755, -163.671, 60.109, 129.834]
  MoveL 222 to (69.42, -37.83, 6.92) mm, rotated rx 90 ry -45.89 rz 90 deg; joints [15.077, -69.53, 129.636, -162.739, 61.234, 125.604]
  MoveL 223 to (68.95, -37.22, 6.38) mm, rotated rx 90 ry -50.05 rz 90 deg; joints [16.009, -68.247, 129.499, -161.879, 62.464, 121.349]
  MoveL 224 to (68.49, -36.58, 5.88) mm, rotated rx 90 ry -54.2 rz 90 deg; joints [16.874, -66.873, 129.353, -161.118, 63.758, 117.196]
  MoveL 225 to (68.02, -35.9, 5.42) mm, rotated rx 90 ry -58.36 rz 90 deg; joints [17.667, -65.415, 129.197, -160.453, 65.105, 113.14]
  MoveL 226 to (67.55, -35.19, 5.02) mm, rotated rx 90 ry -62.52 rz 90 deg; joints [18.386, -63.882, 129.03, -159.882, 66.495, 109.172]
  MoveL 227 to (67.13, -34.29, 4.6) mm, rotated rx 90 ry -67.57 rz 90 deg; joints [19.155, -61.92, 128.8, -159.309, 68.228, 104.454]
  MoveL 228 to (66.72, -33.36, 4.26) mm, rotated rx 90 ry -72.63 rz 90 deg; joints [19.807, -59.872, 128.552, -158.863, 69.997, 99.839]
  MoveL 229 to (66.3, -32.4, 4.01) mm, rotated rx 90 ry -77.68 rz 90 deg; joints [20.339, -57.755, 128.286, -158.537, 71.79, 95.311]
  MoveL 230 to (65.88, -31.42, 3.84) mm, rotated rx 90 ry -82.74 rz 90 deg; joints [20.751, -55.583, 128.002, -158.325, 73.593, 90.855]
  MoveL 231 to (65.46, -30.43, 3.76) mm, rotated rx 90 ry -87.8 rz 90 deg; joints [21.039, -53.372, 127.701, -158.223, 75.397, 86.453]
  MoveL 232 to (65.15, -29.59, 3.75) mm, rotated rx 0 ry -90 rz 180 deg; joints [21.129, -52.375, 127.571, -158.213, 76.211, 84.558]
  MoveL 233 to (64.83, -28.74, 3.75) mm, rotated rx 0 ry -90 rz 180 deg; joints [21.134, -52.326, 127.587, -158.213, 76.273, 84.582]
  MoveL 234 to (64.52, -27.89, 3.75) mm, rotated rx 0 ry -90 rz 180 deg; joints [21.139, -52.277, 127.604, -158.214, 76.334, 84.606]
  MoveL 235 to (64.21, -27.04, 3.75) mm, rotated rx 0 ry -90 rz 180 deg; joints [21.145, -52.227, 127.62, -158.214, 76.396, 84.629]
  MoveL 236 to (63.9, -26.19, 3.75) mm, rotated rx 0 ry -90 rz 180 deg; joints [21.15, -52.178, 127.637, -158.215, 76.458, 84.653]
  MoveL 237 to (63.59, -25.34, 3.75) mm, rotated rx 0 ry -90 rz 180 deg; joints [21.155, -52.128, 127.653, -158.215, 76.519, 84.677]
  MoveL 238 to (61.65, -20.55, 3.75) mm, rotated rx 0 ry -90 rz 180 deg; joints [21.188, -51.853, 127.757, -158.215, 76.875, 84.814]
  MoveL 239 to (59.77, -17.22, 3.75) mm, rotated rx 0 ry -90 rz 180 deg; joints [21.22, -51.675, 127.868, -158.207, 77.146, 84.917]
  MoveL 240 to (57.13, -13.98, 3.75) mm, rotated rx 0 ry -90 rz 180 deg; joints [21.265, -51.524, 128.033, -158.187, 77.443, 85.027]
  MoveL 241 to (55.52, -12.44, 3.75) mm, rotated rx 0 ry -90 rz 180 deg; joints [21.293, -51.462, 128.138, -158.173, 77.6, 85.084]
  MoveL 242 to (53.84, -11.08, 3.75) mm, rotated rx 0 ry -90 rz 180 deg; joints [21.322, -51.414, 128.249, -158.156, 77.751, 85.139]
  MoveL 243 to (52.14, -9.99, 3.75) mm, rotated rx 0 ry -90 rz 180 deg; joints [21.351, -51.384, 128.363, -158.138, 77.887, 85.187]
  MoveL 244 to (50, -9.51, 3.75) mm, rotated rx 0 ry -90 rz 180 deg; joints [21.388, -51.41, 128.515, -158.11, 78.007, 85.227]
  MoveL 245 to (47.86, -9.99, 3.75) mm, rotated rx 0 ry -90 rz 180 deg; joints [21.426, -51.503, 128.676, -158.077, 78.073, 85.245]
  MoveL 246 to (46.16, -11.08, 3.75) mm, rotated rx 0 ry -90 rz 180 deg; joints [21.455, -51.628, 128.811, -158.048, 78.085, 85.243]
  MoveL 247 to (44.48, -12.44, 3.75) mm, rotated rx 0 ry -90 rz 180 deg; joints [21.484, -51.771, 128.946, -158.018, 78.08, 85.234]
  MoveL 248 to (42.87, -13.98, 3.75) mm, rotated rx 0 ry -90 rz 180 deg; joints [21.513, -51.925, 129.078, -157.987, 78.062, 85.219]
  MoveL 249 to (40.23, -17.22, 3.75) mm, rotated rx 0 ry -90 rz 180 deg; joints [21.559, -52.229, 129.3, -157.933, 77.989, 85.178]
  MoveL 250 to (38.35, -20.55, 3.75) mm, rotated rx 0 ry -90 rz 180 deg; joints [21.592, -52.519, 129.466, -157.89, 77.877, 85.123]
  MoveL 251 to (36.41, -25.34, 3.75) mm, rotated rx 0 ry -90 rz 180 deg; joints [21.627, -52.916, 129.647, -157.837, 77.681, 85.033]
  MoveL 252 to (36.1, -26.19, 3.75) mm, rotated rx 0 ry -90 rz 180 deg; joints [21.632, -52.985, 129.677, -157.828, 77.644, 85.016]
  MoveL 253 to (35.79, -27.04, 3.75) mm, rotated rx 0 ry -90 rz 180 deg; joints [21.638, -53.054, 129.706, -157.819, 77.608, 85]
  MoveL 254 to (35.48, -27.89, 3.75) mm, rotated rx 0 ry -90 rz 180 deg; joints [21.643, -53.124, 129.735, -157.81, 77.571, 84.983]
  MoveL 255 to (35.17, -28.74, 3.75) mm, rotated rx 0 ry -90 rz 180 deg; joints [21.649, -53.193, 129.765, -157.801, 77.535, 84.966]
  MoveL 256 to (34.85, -29.59, 3.75) mm, rotated rx 0 ry -90 rz 180 deg; joints [21.654, -53.262, 129.794, -157.792, 77.498, 84.95]
  MoveL 257 to (34.54, -30.43, 3.76) mm, rotated rx 90 ry -87.8 rz 90 deg; joints [21.574, -54.31, 129.973, -157.799, 76.687, 86.835]
  MoveL 258 to (34.12, -31.42, 3.84) mm, rotated rx 90 ry -82.74 rz 90 deg; joints [21.294, -56.62, 130.342, -157.901, 74.861, 91.207]
  MoveL 259 to (33.7, -32.4, 4.01) mm, rotated rx 90 ry -77.68 rz 90 deg; joints [20.888, -58.895, 130.692, -158.114, 73.031, 95.629]
  MoveL 260 to (33.28, -33.36, 4.26) mm, rotated rx 90 ry -72.63 rz 90 deg; joints [20.357, -61.118, 131.024, -158.441, 71.21, 100.119]
  MoveL 261 to (32.87, -34.29, 4.6) mm, rotated rx 90 ry -67.57 rz 90 deg; joints [19.704, -63.274, 131.337, -158.889, 69.408, 104.695]
  MoveL 262 to (32.45, -35.19, 5.02) mm, rotated rx 90 ry -62.52 rz 90 deg; joints [18.93, -65.346, 131.63, -159.465, 67.639, 109.373]
  MoveL 263 to (31.98, -35.9, 5.42) mm, rotated rx 90 ry -58.36 rz 90 deg; joints [18.207, -66.98, 131.867, -160.036, 66.224, 113.308]
  MoveL 264 to (31.51, -36.58, 5.88) mm, rotated rx 90 ry -54.2 rz 90 deg; joints [17.406, -68.54, 132.092, -160.703, 64.85, 117.332]
  MoveL 265 to (31.05, -37.22, 6.38) mm, rotated rx 90 ry -50.05 rz 90 deg; joints [16.53, -70.016, 132.308, -161.467, 63.528, 121.453]
  MoveL 266 to (30.58, -37.83, 6.92) mm, rotated rx 90 ry -45.89 rz 90 deg; joints [15.582, -71.401, 132.513, -162.333, 62.268, 125.677]
  MoveL 267 to (30.04, -38.38, 7.49) mm, rotated rx 90 ry -41.86 rz 90 deg; joints [14.598, -72.654, 132.712, -163.271, 61.118, 129.881]
  MoveL 268 to (29.5, -38.89, 8.1) mm, rotated rx 90 ry -37.83 rz 90 deg; joints [13.553, -73.808, 132.904, -164.308, 60.047, 134.19]
  MoveL 269 to (28.96, -39.35, 8.74) mm, rotated rx 90 ry -33.79 rz 90 deg; joints [12.451, -74.854, 133.091, -165.442, 59.067, 138.605]
  MoveL 270 to (28.42, -39.77, 9.42) mm, rotated rx 90 ry -29.76 rz 90 deg; joints [11.298, -75.788, 133.274, -166.672, 58.19, 143.123]
  MoveL 271 to (27.83, -40.15, 10.15) mm, rotated rx 90 ry -25.52 rz 90 deg; joints [10.034, -76.645, 133.464, -168.062, 57.39, 147.985]
  MoveL 272 to (27.25, -40.48, 10.92) mm, rotated rx 90 ry -21.27 rz 90 deg; joints [8.727, -77.365, 133.651, -169.545, 56.728, 152.949]
  MoveL 273 to (26.67, -40.76, 11.71) mm, rotated rx 90 ry -17.03 rz 90 deg; joints [7.383, -77.943, 133.837, -171.106, 56.215, 158]
  MoveL 274 to (26.08, -40.97, 12.51) mm, rotated rx 90 ry -12.78 rz 90 deg; joints [6.012, -78.374, 134.022, -172.731, 55.862, 163.124]
  MoveL 275 to (25.49, -41.13, 13.34) mm, rotated rx 90 ry -8.49 rz 90 deg; joints [4.605, -78.659, 134.207, -174.421, 55.675, 168.357]
  MoveL 276 to (24.89, -41.22, 14.18) mm, rotated rx 90 ry -4.2 rz 90 deg; joints [3.188, -78.787, 134.392, -176.138, 55.665, 173.622]
  MoveL 277 to (24.3, -41.25, 15.02) mm, rotated rx 90 ry 0 rz 90 deg; joints [1.8, -78.76, 134.571, -177.824, 55.83, 178.777]
  MoveL 278 to (23.7, -41.25, 15.86) mm, rotated rx 90 ry 0 rz 90 deg; joints [1.757, -78.796, 134.617, -177.876, 55.839, 178.807]
  MoveL 279 to (19.04, -41.25, 22.17) mm, rotated rx 90 ry 0 rz 90 deg; joints [1.433, -79.072, 134.971, -178.269, 55.911, 179.03]
  MoveL 280 to (13.72, -41.25, 27.66) mm, rotated rx 90 ry 0 rz 90 deg; joints [1.151, -79.384, 135.369, -178.612, 55.992, 179.224]
  MoveL 281 to (6.48, -41.25, 32.56) mm, rotated rx 90 ry 0 rz 90 deg; joints [0.899, -79.806, 135.903, -178.917, 56.101, 179.396]
  MoveL 282 to (-1.54, -41.25, 36.09) mm, rotated rx 90 ry 0 rz 90 deg; joints [0.716, -80.273, 136.488, -179.138, 56.218, 179.521]
  MoveL 283 to (-9.91, -41.25, 38.42) mm, rotated rx 90 ry 0 rz 90 deg; joints [0.596, -80.762, 137.096, -179.284, 56.336, 179.603]
  MoveL 284 to (-18.44, -41.25, 39.85) mm, rotated rx 90 ry 0 rz 90 deg; joints [0.523, -81.262, 137.711, -179.373, 56.451, 179.653]
  MoveL 285 to (-33.66, -41.25, 41.44) mm, rotated rx 90 ry 0 rz 90 deg; joints [0.443, -82.161, 138.803, -179.47, 56.643, 179.709]
  MoveL 286 to (-37.69, -41.25, 41.93) mm, rotated rx 90 ry 0 rz 90 deg; joints [0.418, -82.401, 139.091, -179.5, 56.691, 179.726]
  MoveL 287 to (-41.59, -41.25, 42.83) mm, rotated rx 90 ry 0 rz 90 deg; joints [0.369, -82.634, 139.369, -179.559, 56.736, 179.758]
  MoveL 288 to (-45.1, -41.25, 44.7) mm, rotated rx 90 ry 0 rz 90 deg; joints [0.266, -82.845, 139.62, -179.683, 56.775, 179.826]
  MoveL 289 to (-50, -41.25, 39.09) mm, rotated rx 90 ry 0 rz 90 deg; joints [0.582, -83.137, 139.965, -179.305, 56.83, 179.62]
  MoveL 290 to (-43.32, -41.25, 37.37) mm, rotated rx 90 ry 0 rz 90 deg; joints [0.674, -82.735, 139.489, -179.195, 56.757, 179.558]
  MoveL 291 to (-36.74, -41.25, 35.17) mm, rotated rx 90 ry 0 rz 90 deg; joints [0.791, -82.34, 139.018, -179.053, 56.682, 179.48]
  MoveL 292 to (-30.12, -41.25, 33.25) mm, rotated rx 90 ry 0 rz 90 deg; joints [0.892, -81.946, 138.544, -178.932, 56.602, 179.412]
  MoveL 293 to (-23.34, -41.25, 32.21) mm, rotated rx 90 ry 0 rz 90 deg; joints [0.943, -81.544, 138.057, -178.87, 56.517, 179.376]
  MoveL 294 to (-16.33, -41.25, 31.5) mm, rotated rx 90 ry 0 rz 90 deg; joints [0.975, -81.132, 137.552, -178.829, 56.426, 179.353]
  MoveL 295 to (-9.37, -41.25, 30.15) mm, rotated rx 90 ry 0 rz 90 deg; joints [1.042, -80.723, 137.048, -178.748, 56.331, 179.306]
  MoveL 296 to (-2.68, -41.25, 27.82) mm, rotated rx 90 ry 0 rz 90 deg; joints [1.16, -80.332, 136.561, -178.605, 56.238, 179.224]
  MoveL 297 to (3.46, -41.25, 24.48) mm, rotated rx 90 ry 0 rz 90 deg; joints [1.331, -79.972, 136.111, -178.397, 56.15, 179.107]
  MoveL 298 to (8.93, -41.25, 20.18) mm, rotated rx 90 ry 0 rz 90 deg; joints [1.553, -79.65, 135.705, -178.129, 56.069, 178.955]
  MoveL 299 to (11.76, -41.25, 17.39) mm, rotated rx 90 ry 0 rz 90 deg; joints [1.696, -79.483, 135.493, -177.955, 56.028, 178.857]
  MoveL 300 to (12.43, -41.25, 16.64) mm, rotated rx 90 ry 0 rz 90 deg; joints [1.735, -79.442, 135.443, -177.908, 56.018, 178.83]
  MoveL 301 to (13.1, -41.25, 15.88) mm, rotated rx 90 ry 0 rz 90 deg; joints [1.774, -79.402, 135.392, -177.861, 56.008, 178.804]
  MoveL 302 to (13.78, -41.25, 15.12) mm, rotated rx 90 ry 0 rz 90 deg; joints [1.812, -79.362, 135.341, -177.814, 55.998, 178.777]
  MoveL 303 to (14.45, -41.23, 14.36) mm, rotated rx 90 ry -3.25 rz 90 deg; joints [2.903, -79.384, 135.186, -176.491, 55.851, 174.775]
  MoveL 304 to (15.09, -41.16, 13.55) mm, rotated rx 90 ry -7.41 rz 90 deg; joints [4.289, -79.291, 135.002, -174.813, 55.82, 169.67]
  MoveL 305 to (15.73, -41.02, 12.74) mm, rotated rx 90 ry -11.57 rz 90 deg; joints [5.668, -79.049, 134.818, -173.155, 55.959, 164.587]
  MoveL 306 to (16.38, -40.83, 11.95) mm, rotated rx 90 ry -15.73 rz 90 deg; joints [7.03, -78.661, 134.632, -171.537, 56.262, 159.55]
  MoveL 307 to (17.02, -40.58, 11.17) mm, rotated rx 90 ry -19.88 rz 90 deg; joints [8.367, -78.129, 134.445, -169.977, 56.722, 154.578]
  MoveL 308 to (17.6, -40.28, 10.43) mm, rotated rx 90 ry -23.97 rz 90 deg; joints [9.65, -77.473, 134.264, -168.512, 57.32, 149.765]
  MoveL 309 to (18.18, -39.93, 9.71) mm, rotated rx 90 ry -28.06 rz 90 deg; joints [10.895, -76.687, 134.081, -167.129, 58.052, 145.044]
  MoveL 310 to (18.76, -39.52, 9.01) mm, rotated rx 90 ry -32.15 rz 90 deg; joints [12.094, -75.776, 133.895, -165.838, 58.906, 140.424]
  MoveL 311 to (19.34, -39.07, 8.35) mm, rotated rx 90 ry -36.24 rz 90 deg; joints [13.242, -74.746, 133.705, -164.643, 59.872, 135.91]
  MoveL 312 to (19.84, -38.58, 7.73) mm, rotated rx 90 ry -40.29 rz 90 deg; joints [14.322, -73.62, 133.519, -163.559, 60.926, 131.554]
  MoveL 313 to (20.33, -38.05, 7.14) mm, rotated rx 90 ry -44.33 rz 90 deg; joints [15.342, -72.39, 133.326, -162.574, 62.065, 127.306]
  MoveL 314 to (20.82, -37.47, 6.59) mm, rotated rx 90 ry -48.37 rz 90 deg; joints [16.297, -71.062, 133.127, -161.689, 63.279, 123.162]
  MoveL 315 to (21.32, -36.86, 6.08) mm, rotated rx 90 ry -52.42 rz 90 deg; joints [17.185, -69.644, 132.918, -160.901, 64.556, 119.12]
  MoveL 316 to (21.73, -36.14, 5.58) mm, rotated rx 90 ry -56.9 rz 90 deg; joints [18.088, -67.982, 132.687, -160.137, 66.035, 114.755]
  MoveL 317 to (22.14, -35.39, 5.12) mm, rotated rx 90 ry -61.38 rz 90 deg; joints [18.901, -66.229, 132.442, -159.485, 67.568, 110.497]
  MoveL 318 to (22.55, -34.6, 4.73) mm, rotated rx 90 ry -65.86 rz 90 deg; joints [19.621, -64.394, 132.183, -158.939, 69.141, 106.337]
  MoveL 319 to (22.97, -33.79, 4.41) mm, rotated rx 90 ry -70.34 rz 90 deg; joints [20.247, -62.489, 131.91, -158.495, 70.744, 102.261]
  MoveL 320 to (23.34, -32.85, 4.12) mm, rotated rx 90 ry -75.32 rz 90 deg; joints [20.831, -60.304, 131.593, -158.114, 72.553, 97.811]
  MoveL 321 to (23.72, -31.89, 3.91) mm, rotated rx 90 ry -80.31 rz 90 deg; joints [21.293, -58.061, 131.258, -157.848, 74.375, 93.437]
  MoveL 322 to (24.09, -30.92, 3.79) mm, rotated rx 90 ry -85.29 rz 90 deg; joints [21.633, -55.775, 130.904, -157.69, 76.198, 89.119]
  MoveL 323 to (24.46, -29.95, 3.75) mm, rotated rx 0 ry -90 rz 180 deg; joints [21.84, -53.585, 130.552, -157.638, 77.916, 85.078]
  MoveL 324 to (26.01, -26.09, 3.75) mm, rotated rx 0 ry -90 rz 180 deg; joints [21.813, -53.264, 130.41, -157.681, 78.079, 85.153]
  MoveL 325 to (29.8, -19.01, 3.75) mm, rotated rx 0 ry -90 rz 180 deg; joints [21.744, -52.649, 130.075, -157.773, 78.334, 85.276]
  MoveL 326 to (34.48, -12.81, 3.75) mm, rotated rx 0 ry -90 rz 180 deg; joints [21.661, -52.074, 129.679, -157.871, 78.493, 85.362]
  MoveL 327 to (39.73, -7.1, 3.75) mm, rotated rx 0 ry -90 rz 180 deg; joints [21.568, -51.522, 129.242, -157.975, 78.593, 85.425]
  MoveL 328 to (45.25, -1.49, 3.75) mm, rotated rx 0 ry -90 rz 180 deg; joints [21.471, -50.971, 128.784, -158.08, 78.67, 85.48]
  MoveL 329 to (54.75, -1.49, 3.75) mm, rotated rx 0 ry -90 rz 180 deg; joints [21.306, -50.713, 128.089, -158.215, 78.252, 85.348]
  MoveL 330 to (60.27, -7.1, 3.75) mm, rotated rx 0 ry -90 rz 180 deg; joints [21.212, -50.954, 127.738, -158.264, 77.694, 85.143]
  MoveL 331 to (65.52, -12.81, 3.75) mm, rotated rx 0 ry -90 rz 180 deg; joints [21.122, -51.203, 127.404, -158.307, 77.144, 84.942]
  MoveL 332 to (70.2, -19.01, 3.75) mm, rotated rx 0 ry -90 rz 180 deg; joints [21.043, -51.497, 127.112, -158.338, 76.592, 84.738]
  MoveL 333 to (73.99, -26.09, 3.75) mm, rotated rx 0 ry -90 rz 180 deg; joints [20.98, -51.872, 126.888, -158.349, 76.03, 84.526]
  MoveL 334 to (75.53, -29.95, 3.75) mm, rotated rx 0 ry -90 rz 180 deg; joints [20.954, -52.089, 126.803, -158.347, 75.747, 84.418]
  MoveL 335 to (75.91, -30.92, 3.79) mm, rotated rx 90 ry -85.29 rz 90 deg; joints [20.741, -54.143, 127.091, -158.392, 74.083, 88.51]
  MoveL 336 to (76.28, -31.89, 3.91) mm, rotated rx 90 ry -80.31 rz 90 deg; joints [20.4, -56.285, 127.381, -158.54, 72.322, 92.888]
  MoveL 337 to (76.66, -32.85, 4.12) mm, rotated rx 90 ry -75.32 rz 90 deg; joints [19.941, -58.381, 127.654, -158.798, 70.567, 97.325]
  MoveL 338 to (77.03, -33.79, 4.41) mm, rotated rx 90 ry -70.34 rz 90 deg; joints [19.366, -60.419, 127.91, -159.169, 68.828, 101.84]
  MoveL 339 to (77.44, -34.6, 4.73) mm, rotated rx 90 ry -65.86 rz 90 deg; joints [18.751, -62.184, 128.119, -159.605, 67.286, 105.974]
  MoveL 340 to (77.86, -35.39, 5.12) mm, rotated rx 90 ry -61.38 rz 90 deg; joints [18.046, -63.879, 128.315, -160.142, 65.777, 110.194]
  MoveL 341 to (78.27, -36.14, 5.58) mm, rotated rx 90 ry -56.9 rz 90 deg; joints [17.253, -65.493, 128.497, -160.785, 64.31, 114.511]
  MoveL 342 to (78.68, -36.86, 6.08) mm, rotated rx 90 ry -52.42 rz 90 deg; joints [16.375, -67.017, 128.668, -161.536, 62.898, 118.933]
  MoveL 343 to (79.17, -37.47, 6.59) mm, rotated rx 90 ry -48.37 rz 90 deg; joints [15.512, -68.301, 128.803, -162.313, 61.676, 123.022]
  MoveL 344 to (79.67, -38.05, 7.14) mm, rotated rx 90 ry -44.33 rz 90 deg; joints [14.585, -69.498, 128.931, -163.185, 60.517, 127.211]
  MoveL 345 to (80.16, -38.58, 7.73) mm, rotated rx 90 ry -40.29 rz 90 deg; joints [13.6, -70.6, 129.051, -164.151, 59.432, 131.5]
  MoveL 346 to (80.66, -39.07, 8.35) mm, rotated rx 90 ry -36.24 rz 90 deg; joints [12.56, -71.601, 129.166, -165.213, 58.432, 135.891]
  MoveL 347 to (81.24, -39.52, 9.01) mm, rotated rx 90 ry -32.15 rz 90 deg; joints [11.456, -72.502, 129.271, -166.381, 57.514, 140.435]
  MoveL 348 to (81.82, -39.93, 9.71) mm, rotated rx 90 ry -28.06 rz 90 deg; joints [10.307, -73.288, 129.372, -167.639, 56.703, 145.078]
  MoveL 349 to (82.4, -40.28, 10.43) mm, rotated rx 90 ry -23.97 rz 90 deg; joints [9.118, -73.956, 129.469, -168.982, 56.009, 149.814]
  MoveL 350 to (82.98, -40.58, 11.17) mm, rotated rx 90 ry -19.88 rz 90 deg; joints [7.895, -74.501, 129.565, -170.399, 55.442, 154.636]
  MoveL 351 to (83.62, -40.83, 11.95) mm, rotated rx 90 ry -15.73 rz 90 deg; joints [6.624, -74.924, 129.655, -171.905, 55.002, 159.61]
  MoveL 352 to (84.27, -41.02, 12.74) mm, rotated rx 90 ry -11.57 rz 90 deg; joints [5.334, -75.212, 129.744, -173.461, 54.709, 164.642]
  MoveL 353 to (84.91, -41.16, 13.55) mm, rotated rx 90 ry -7.41 rz 90 deg; joints [4.031, -75.364, 129.831, -175.05, 54.568, 169.715]
  MoveL 354 to (85.55, -41.23, 14.36) mm, rotated rx 90 ry -3.25 rz 90 deg; joints [2.725, -75.379, 129.915, -176.656, 54.582, 174.806]
  MoveL 355 to (86.22, -41.25, 15.12) mm, rotated rx 90 ry 0 rz 90 deg; joints [1.699, -75.285, 129.966, -177.918, 54.698, 178.796]
  MoveL 356 to (86.9, -41.25, 15.88) mm, rotated rx 90 ry 0 rz 90 deg; joints [1.661, -75.249, 129.916, -177.965, 54.684, 178.823]
  MoveL 357 to (87.57, -41.25, 16.64) mm, rotated rx 90 ry 0 rz 90 deg; joints [1.622, -75.213, 129.867, -178.011, 54.67, 178.85]
  MoveL 358 to (88.25, -41.25, 17.39) mm, rotated rx 90 ry 0 rz 90 deg; joints [1.584, -75.177, 129.818, -178.058, 54.656, 178.876]
  MoveL 359 to (91.07, -41.25, 20.18) mm, rotated rx 90 ry 0 rz 90 deg; joints [1.443, -75.025, 129.61, -178.23, 54.598, 178.974]
  MoveL 360 to (96.54, -41.25, 24.48) mm, rotated rx 90 ry 0 rz 90 deg; joints [1.225, -74.729, 129.203, -178.495, 54.483, 179.126]
  MoveL 361 to (102.68, -41.25, 27.82) mm, rotated rx 90 ry 0 rz 90 deg; joints [1.056, -74.394, 128.741, -178.701, 54.354, 179.243]
  MoveL 362 to (109.37, -41.25, 30.15) mm, rotated rx 90 ry 0 rz 90 deg; joints [0.937, -74.029, 128.235, -178.845, 54.211, 179.324]
  MoveL 363 to (116.33, -41.25, 31.5) mm, rotated rx 90 ry 0 rz 90 deg; joints [0.866, -73.649, 127.704, -178.93, 54.06, 179.372]
  MoveL 364 to (123.34, -41.25, 32.21) mm, rotated rx 90 ry 0 rz 90 deg; joints [0.827, -73.266, 127.167, -178.976, 53.905, 179.397]
  MoveL 365 to (130.13, -41.25, 33.25) mm, rotated rx 90 ry 0 rz 90 deg; joints [0.773, -72.897, 126.646, -179.042, 53.752, 179.433]
  MoveL 366 to (136.74, -41.25, 35.17) mm, rotated rx 90 ry 0 rz 90 deg; joints [0.678, -72.538, 126.137, -179.158, 53.601, 179.5]
  MoveL 367 to (143.32, -41.25, 37.37) mm, rotated rx 90 ry 0 rz 90 deg; joints [0.57, -72.183, 125.629, -179.29, 53.449, 179.577]
  MoveL 368 to (150, -41.25, 39.09) mm, rotated rx 90 ry 0 rz 90 deg; joints [0.487, -71.821, 125.11, -179.393, 53.291, 179.637]
  MoveL 369 to (150, -41.25, 31.96) mm, rotated rx 90 ry 0 rz 90 deg; joints [0.821, -71.816, 125.104, -178.976, 53.292, 179.388]
  MoveL 370 to (144.93, -41.25, 28.57) mm, rotated rx 90 ry 0 rz 90 deg; joints [0.984, -72.088, 125.494, -178.774, 53.412, 179.269]
  MoveL 371 to (139.35, -41.25, 26.34) mm, rotated rx 90 ry 0 rz 90 deg; joints [1.094, -72.389, 125.924, -178.64, 53.543, 179.192]
  MoveL 372 to (133.44, -41.25, 24.88) mm, rotated rx 90 ry 0 rz 90 deg; joints [1.169, -72.709, 126.379, -178.55, 53.679, 179.141]
  MoveL 373 to (127.36, -41.25, 23.82) mm, rotated rx 90 ry 0 rz 90 deg; joints [1.226, -73.039, 126.847, -178.482, 53.817, 179.103]
  MoveL 374 to (121.16, -41.25, 22.72) mm, rotated rx 90 ry 0 rz 90 deg; joints [1.284, -73.376, 127.322, -178.411, 53.956, 179.065]
  MoveL 375 to (115.12, -41.25, 21.22) mm, rotated rx 90 ry 0 rz 90 deg; joints [1.363, -73.704, 127.781, -178.316, 54.089, 179.012]
  MoveL 376 to (109.45, -41.25, 18.9) mm, rotated rx 90 ry 0 rz 90 deg; joints [1.482, -74.012, 128.211, -178.173, 54.212, 178.931]
  MoveL 377 to (104.25, -41.25, 15.52) mm, rotated rx 90 ry 0 rz 90 deg; joints [1.654, -74.292, 128.6, -177.964, 54.325, 178.812]
  MoveL 378 to (103.32, -41.24, 14.62) mm, rotated rx 90 ry -1.91 rz 90 deg; joints [2.269, -74.386, 128.611, -177.204, 54.258, 176.454]
  MoveL 379 to (102.38, -41.18, 13.74) mm, rotated rx 90 ry -6.45 rz 90 deg; joints [3.675, -74.424, 128.54, -175.467, 54.201, 170.893]
  MoveL 380 to (101.44, -41.04, 12.86) mm, rotated rx 90 ry -10.99 rz 90 deg; joints [5.079, -74.302, 128.465, -173.744, 54.325, 165.35]
  MoveL 381 to (100.5, -40.84, 11.99) mm, rotated rx 90 ry -15.53 rz 90 deg; joints [6.471, -74.02, 128.387, -172.056, 54.629, 159.85]
  MoveL 382 to (99.57, -40.57, 11.14) mm, rotated rx 90 ry -20.07 rz 90 deg; joints [7.841, -73.581, 128.307, -170.426, 55.103, 154.416]
  MoveL 383 to (98.79, -40.21, 10.27) mm, rotated rx 90 ry -24.87 rz 90 deg; joints [9.251, -72.941, 128.203, -168.789, 55.777, 148.774]
  MoveL 384 to (98.01, -39.78, 9.43) mm, rotated rx 90 ry -29.66 rz 90 deg; joints [10.614, -72.136, 128.095, -167.257, 56.619, 143.247]
  MoveL 385 to (97.23, -39.28, 8.63) mm, rotated rx 90 ry -34.45 rz 90 deg; joints [11.92, -71.172, 127.981, -165.842, 57.614, 137.851]
  MoveL 386 to (96.45, -38.71, 7.88) mm, rotated rx 90 ry -39.25 rz 90 deg; joints [13.161, -70.059, 127.862, -164.554, 58.746, 132.592]
  MoveL 387 to (95.77, -38.09, 7.18) mm, rotated rx 90 ry -44.05 rz 90 deg; joints [14.329, -68.797, 127.727, -163.395, 59.999, 127.466]
  MoveL 388 to (95.08, -37.4, 6.53) mm, rotated rx 90 ry -48.86 rz 90 deg; joints [15.415, -67.403, 127.583, -162.37, 61.355, 122.482]
  MoveL 389 to (94.39, -36.67, 5.94) mm, rotated rx 90 ry -53.66 rz 90 deg; joints [16.413, -65.887, 127.428, -161.476, 62.8, 117.632]
  MoveL 390 to (93.71, -35.88, 5.41) mm, rotated rx 90 ry -58.46 rz 90 deg; joints [17.32, -64.26, 127.26, -160.711, 64.317, 112.911]
  MoveL 391 to (93.12, -35.05, 4.95) mm, rotated rx 90 ry -63.33 rz 90 deg; joints [18.136, -62.507, 127.068, -160.063, 65.907, 108.252]
  MoveL 392 to (92.53, -34.18, 4.55) mm, rotated rx 90 ry -68.19 rz 90 deg; joints [18.85, -60.666, 126.86, -159.537, 67.544, 103.699]
  MoveL 393 to (91.94, -33.28, 4.24) mm, rotated rx 90 ry -73.05 rz 90 deg; joints [19.457, -58.748, 126.637, -159.127, 69.212, 99.242]
  MoveL 394 to (91.35, -32.36, 4) mm, rotated rx 90 ry -77.91 rz 90 deg; joints [19.956, -56.767, 126.397, -158.827, 70.902, 94.864]
  MoveL 395 to (90.92, -31.56, 3.86) mm, rotated rx 90 ry -82.03 rz 90 deg; joints [20.292, -55.046, 126.175, -158.657, 72.34, 91.205]
  MoveL 396 to (90.5, -30.75, 3.77) mm, rotated rx 90 ry -86.16 rz 90 deg; joints [20.548, -53.297, 125.942, -158.559, 73.781, 87.582]
  MoveL 397 to (90.07, -29.95, 3.75) mm, rotated rx 0 ry -90 rz 180 deg; joints [20.714, -51.647, 125.717, -158.533, 75.125, 84.235]
  MoveL 398 to (89.65, -29.14, 3.75) mm, rotated rx 0 ry -90 rz 180 deg; joints [20.721, -51.606, 125.743, -158.532, 75.188, 84.259]
  MoveL 399 to (89.22, -28.33, 3.75) mm, rotated rx 0 ry -90 rz 180 deg; joints [20.728, -51.564, 125.769, -158.531, 75.252, 84.283]
  MoveL 400 to (87.07, -24.08, 3.75) mm, rotated rx 0 ry -90 rz 180 deg; joints [20.763, -51.343, 125.897, -158.528, 75.58, 84.406]
  MoveL 401 to (84.65, -19.99, 3.75) mm, rotated rx 0 ry -90 rz 180 deg; joints [20.803, -51.138, 126.045, -158.52, 75.912, 84.529]
  MoveL 402 to (80.12, -14.74, 3.75) mm, rotated rx 0 ry -90 rz 180 deg; joints [20.878, -50.914, 126.338, -158.49, 76.4, 84.706]
  MoveL 403 to (74.83, -10.27, 3.75) mm, rotated rx 0 ry -90 rz 180 deg; joints [20.966, -50.761, 126.691, -158.444, 76.879, 84.876]
  MoveL 404 to (69.43, -5.9, 3.75) mm, rotated rx 0 ry -90 rz 180 deg; joints [21.056, -50.613, 127.05, -158.395, 77.358, 85.046]
  MoveL 405 to (64.56, -1, 3.75) mm, rotated rx 0 ry -90 rz 180 deg; joints [21.139, -50.408, 127.362, -158.352, 77.846, 85.223]
  MoveL 406 to (35.45, -1, 3.75) mm, rotated rx 0 ry -90 rz 180 deg; joints [21.644, -51.2, 129.493, -157.94, 79.129, 85.63]
  MoveL 407 to (30.57, -5.9, 3.75) mm, rotated rx 0 ry -90 rz 180 deg; joints [21.731, -51.683, 129.897, -157.846, 79.062, 85.582]
  MoveL 408 to (25.17, -10.27, 3.75) mm, rotated rx 0 ry -90 rz 180 deg; joints [21.828, -52.144, 130.331, -157.746, 79.044, 85.553]
  MoveL 409 to (19.88, -14.74, 3.75) mm, rotated rx 0 ry -90 rz 180 deg; joints [21.923, -52.612, 130.755, -157.645, 79.011, 85.518]
  MoveL 410 to (15.35, -19.99, 3.75) mm, rotated rx 0 ry -90 rz 180 deg; joints [22.006, -53.118, 131.129, -157.551, 78.895, 85.45]
  MoveL 411 to (12.93, -24.08, 3.75) mm, rotated rx 0 ry -90 rz 180 deg; joints [22.05, -53.484, 131.338, -157.495, 78.755, 85.381]
  MoveL 412 to (10.78, -28.33, 3.75) mm, rotated rx 0 ry -90 rz 180 deg; joints [22.09, -53.853, 131.527, -157.44, 78.591, 85.302]
  MoveL 413 to (10.35, -29.14, 3.75) mm, rotated rx 0 ry -90 rz 180 deg; joints [22.098, -53.924, 131.564, -157.43, 78.561, 85.287]
  MoveL 414 to (9.93, -29.95, 3.75) mm, rotated rx 0 ry -90 rz 180 deg; joints [22.106, -53.995, 131.601, -157.419, 78.53, 85.272]
  MoveL 415 to (9.5, -30.75, 3.77) mm, rotated rx 90 ry -86.16 rz 90 deg; joints [21.946, -55.814, 131.901, -157.457, 77.113, 88.552]
  MoveL 416 to (9.08, -31.56, 3.86) mm, rotated rx 90 ry -82.03 rz 90 deg; joints [21.691, -57.746, 132.208, -157.567, 75.587, 92.098]
  MoveL 417 to (8.65, -32.36, 4) mm, rotated rx 90 ry -77.91 rz 90 deg; joints [21.351, -59.652, 132.502, -157.751, 74.06, 95.677]
  MoveL 418 to (8.06, -33.28, 4.24) mm, rotated rx 90 ry -73.05 rz 90 deg; joints [20.843, -61.859, 132.839, -158.065, 72.267, 99.956]
  MoveL 419 to (7.47, -34.18, 4.55) mm, rotated rx 90 ry -68.19 rz 90 deg; joints [20.219, -64.005, 133.156, -158.49, 70.49, 104.313]
  MoveL 420 to (6.88, -35.05, 4.95) mm, rotated rx 90 ry -63.33 rz 90 deg; joints [19.481, -66.075, 133.456, -159.032, 68.741, 108.764]
  MoveL 421 to (6.29, -35.88, 5.41) mm, rotated rx 90 ry -58.46 rz 90 deg; joints [18.631, -68.054, 133.738, -159.698, 67.034, 113.322]
  MoveL 422 to (5.61, -36.67, 5.94) mm, rotated rx 90 ry -53.66 rz 90 deg; joints [17.685, -69.911, 134.009, -160.482, 65.405, 117.948]
  MoveL 423 to (4.92, -37.4, 6.53) mm, rotated rx 90 ry -48.86 rz 90 deg; joints [16.637, -71.654, 134.265, -161.4, 63.847, 122.706]
  MoveL 424 to (4.23, -38.09, 7.18) mm, rotated rx 90 ry -44.05 rz 90 deg; joints [15.491, -73.268, 134.509, -162.455, 62.377, 127.608]
  MoveL 425 to (3.55, -38.71, 7.88) mm, rotated rx 90 ry -39.25 rz 90 deg; joints [14.253, -74.743, 134.743, -163.652, 61.014, 132.661]
  MoveL 426 to (2.77, -39.28, 8.63) mm, rotated rx 90 ry -34.45 rz 90 deg; joints [12.934, -76.068, 134.975, -164.987, 59.78, 137.858]
  MoveL 427 to (1.99, -39.78, 9.43) mm, rotated rx 90 ry -29.66 rz 90 deg; joints [11.539, -77.231, 135.201, -166.46, 58.692, 143.207]
  MoveL 428 to (1.21, -40.21, 10.27) mm, rotated rx 90 ry -24.87 rz 90 deg; joints [10.075, -78.222, 135.423, -168.064, 57.768, 148.702]
  MoveL 429 to (0.43, -40.57, 11.14) mm, rotated rx 90 ry -20.07 rz 90 deg; joints [8.555, -79.033, 135.642, -169.786, 57.028, 154.327]
  MoveL 430 to (-0.5, -40.84, 11.99) mm, rotated rx 90 ry -15.53 rz 90 deg; joints [7.075, -79.639, 135.863, -171.507, 56.515, 159.758]
  MoveL 431 to (-1.44, -41.04, 12.86) mm, rotated rx 90 ry -10.99 rz 90 deg; joints [5.564, -80.072, 136.083, -173.299, 56.193, 165.268]
  MoveL 432 to (-2.38, -41.18, 13.74) mm, rotated rx 90 ry -6.45 rz 90 deg; joints [4.034, -80.325, 136.302, -175.137, 56.073, 170.829]
  MoveL 433 to (-3.32, -41.24, 14.62) mm, rotated rx 90 ry -1.91 rz 90 deg; joints [2.496, -80.397, 136.52, -176.995, 56.16, 176.413]
  MoveL 434 to (-4.25, -41.25, 15.52) mm, rotated rx 90 ry 0 rz 90 deg; joints [1.822, -80.404, 136.652, -177.809, 56.267, 178.783]
  MoveL 435 to (-9.45, -41.25, 18.9) mm, rotated rx 90 ry 0 rz 90 deg; joints [1.648, -80.712, 137.035, -178.02, 56.338, 178.902]
  MoveL 436 to (-15.12, -41.25, 21.22) mm, rotated rx 90 ry 0 rz 90 deg; joints [1.532, -81.048, 137.449, -178.162, 56.415, 178.983]
  MoveL 437 to (-21.16, -41.25, 22.72) mm, rotated rx 90 ry 0 rz 90 deg; joints [1.458, -81.404, 137.885, -178.251, 56.494, 179.034]
  MoveL 438 to (-27.36, -41.25, 23.82) mm, rotated rx 90 ry 0 rz 90 deg; joints [1.407, -81.771, 138.332, -178.314, 56.572, 179.071]
  MoveL 439 to (-33.44, -41.25, 24.88) mm, rotated rx 90 ry 0 rz 90 deg; joints [1.356, -82.133, 138.769, -178.376, 56.647, 179.107]
  MoveL 440 to (-39.35, -41.25, 26.34) mm, rotated rx 90 ry 0 rz 90 deg; joints [1.283, -82.487, 139.193, -178.465, 56.716, 179.157]
  MoveL 441 to (-44.93, -41.25, 28.57) mm, rotated rx 90 ry 0 rz 90 deg; joints [1.166, -82.823, 139.593, -178.606, 56.778, 179.236]
  MoveL 442 to (-50, -41.25, 31.96) mm, rotated rx 90 ry 0 rz 90 deg; joints [0.981, -83.131, 139.958, -178.828, 56.832, 179.359]
  MoveL 443 to (-50, -41.25, 30.97) mm, rotated rx 90 ry 0 rz 90 deg; joints [1.037, -83.13, 139.956, -178.761, 56.833, 179.322]
  MoveL 444 to (-50, -41.25, 29.97) mm, rotated rx 90 ry 0 rz 90 deg; joints [1.093, -83.129, 139.955, -178.694, 56.833, 179.286]
  MoveL 445 to (-50, -41.25, 28.98) mm, rotated rx 90 ry 0 rz 90 deg; joints [1.149, -83.128, 139.954, -178.628, 56.834, 179.249]
  MoveL 446 to (-50, -41.25, 27.98) mm, rotated rx 90 ry 0 rz 90 deg; joints [1.205, -83.126, 139.952, -178.561, 56.834, 179.213]
  MoveL 447 to (-50, -41.25, 26.99) mm, rotated rx 90 ry 0 rz 90 deg; joints [1.26, -83.125, 139.951, -178.494, 56.835, 179.176]
  MoveL 448 to (-50, -41.25, 25.99) mm, rotated rx 90 ry 0 rz 90 deg; joints [1.316, -83.124, 139.949, -178.428, 56.835, 179.14]
  MoveL 449 to (-50, -41.25, 25) mm, rotated rx 90 ry 0 rz 90 deg; joints [1.372, -83.122, 139.948, -178.361, 56.836, 179.103]
  MoveL 450 to (-50, -41.25, 24) mm, rotated rx 90 ry 0 rz 90 deg; joints [1.428, -83.121, 139.946, -178.294, 56.837, 179.067]
  MoveL 451 to (-50, -41.25, 23.01) mm, rotated rx 90 ry 0 rz 90 deg; joints [1.483, -83.119, 139.944, -178.228, 56.837, 179.03]
  MoveL 452 to (-50, -41.25, 22.01) mm, rotated rx 90 ry 0 rz 90 deg; joints [1.539, -83.118, 139.942, -178.161, 56.838, 178.994]
  MoveL 453 to (-50, -41.25, 21.02) mm, rotated rx 90 ry 0 rz 90 deg; joints [1.595, -83.116, 139.94, -178.095, 56.839, 178.957]
  MoveL 454 to (-50, -41.25, 20.02) mm, rotated rx 90 ry 0 rz 90 deg; joints [1.651, -83.114, 139.938, -178.028, 56.839, 178.921]
  MoveL 455 to (-50, -41.25, 19.03) mm, rotated rx 90 ry 0 rz 90 deg; joints [1.707, -83.113, 139.936, -177.961, 56.84, 178.885]
  MoveL 456 to (-50, -41.25, 18.03) mm, rotated rx 90 ry 0 rz 90 deg; joints [1.762, -83.111, 139.934, -177.895, 56.841, 178.848]
  MoveL 457 to (-50, -41.25, 17.04) mm, rotated rx 90 ry 0 rz 90 deg; joints [1.818, -83.109, 139.932, -177.828, 56.842, 178.812]
  MoveL 458 to (-50, -41.25, 16.04) mm, rotated rx 90 ry 0 rz 90 deg; joints [1.874, -83.107, 139.93, -177.762, 56.843, 178.775]
  MoveL 459 to (-50, -41.25, 15.05) mm, rotated rx 90 ry 0 rz 90 deg; joints [1.93, -83.105, 139.927, -177.695, 56.843, 178.739]
  MoveL 460 to (-50, -41.21, 14.05) mm, rotated rx 90 ry -4.83 rz 90 deg; joints [3.647, -83.164, 139.763, -175.635, 56.675, 172.765]
  MoveL 461 to (-50, -41.08, 13.07) mm, rotated rx 90 ry -9.9 rz 90 deg; joints [5.442, -82.989, 139.59, -173.49, 56.772, 166.521]
  MoveL 462 to (-50, -40.87, 12.09) mm, rotated rx 90 ry -14.97 rz 90 deg; joints [7.219, -82.574, 139.418, -171.396, 57.14, 160.337]
  MoveL 463 to (-50, -40.57, 11.14) mm, rotated rx 90 ry -20.04 rz 90 deg; joints [8.96, -81.927, 139.246, -169.391, 57.767, 154.257]
  MoveL 464 to (-49.08, -40.7, 11.54) mm, rotated rx 90 ry -17.93 rz 90 deg; joints [8.236, -82.17, 139.253, -170.218, 57.465, 156.767]
  MoveL 465 to (-48.17, -40.82, 11.93) mm, rotated rx 90 ry -15.83 rz 90 deg; joints [7.505, -82.372, 139.259, -171.062, 57.207, 159.299]
  MoveL 466 to (-47.25, -40.93, 12.33) mm, rotated rx 90 ry -13.73 rz 90 deg; joints [6.769, -82.534, 139.266, -171.92, 56.993, 161.849]
  MoveL 467 to (-46.33, -41.02, 12.73) mm, rotated rx 90 ry -11.63 rz 90 deg; joints [6.029, -82.656, 139.272, -172.791, 56.825, 164.414]
  MoveL 468 to (-45.37, -41.06, 12.93) mm, rotated rx 90 ry -10.62 rz 90 deg; joints [5.669, -82.668, 139.238, -173.217, 56.755, 165.653]
  MoveL 469 to (-44.41, -41.09, 13.12) mm, rotated rx 90 ry -9.61 rz 90 deg; joints [5.309, -82.672, 139.205, -173.643, 56.695, 166.894]
  MoveL 470 to (-43.45, -41.12, 13.32) mm, rotated rx 90 ry -8.6 rz 90 deg; joints [4.949, -82.665, 139.171, -174.072, 56.647, 168.138]
  MoveL 471 to (-42.49, -41.15, 13.52) mm, rotated rx 90 ry -7.59 rz 90 deg; joints [4.589, -82.649, 139.137, -174.501, 56.609, 169.382]
  MoveL 472 to (-41.5, -41.15, 13.51) mm, rotated rx 90 ry -7.62 rz 90 deg; joints [4.598, -82.589, 139.066, -174.489, 56.599, 169.337]
  MoveL 473 to (-40.52, -41.15, 13.5) mm, rotated rx 90 ry -7.66 rz 90 deg; joints [4.607, -82.529, 138.995, -174.478, 56.588, 169.292]
  MoveL 474 to (-39.54, -41.15, 13.49) mm, rotated rx 90 ry -7.7 rz 90 deg; joints [4.616, -82.469, 138.924, -174.466, 56.578, 169.246]
  MoveL 475 to (-38.56, -41.15, 13.48) mm, rotated rx 90 ry -7.74 rz 90 deg; joints [4.626, -82.409, 138.853, -174.454, 56.567, 169.2]
  MoveL 476 to (-37.58, -41.12, 13.28) mm, rotated rx 90 ry -8.78 rz 90 deg; joints [4.984, -82.308, 138.748, -174.025, 56.584, 167.925]
  MoveL 477 to (-36.6, -41.09, 13.08) mm, rotated rx 90 ry -9.81 rz 90 deg; joints [5.342, -82.196, 138.643, -173.598, 56.612, 166.653]
  MoveL 478 to (-35.62, -41.05, 12.88) mm, rotated rx 90 ry -10.85 rz 90 deg; joints [5.698, -82.075, 138.538, -173.173, 56.651, 165.382]
  MoveL 479 to (-34.64, -41.01, 12.68) mm, rotated rx 90 ry -11.89 rz 90 deg; joints [6.053, -81.944, 138.434, -172.752, 56.701, 164.115]
  MoveL 480 to (-33.66, -40.97, 12.48) mm, rotated rx 90 ry -12.93 rz 90 deg; joints [6.406, -81.804, 138.329, -172.334, 56.761, 162.851]
  MoveL 481 to (-32.68, -40.92, 12.28) mm, rotated rx 90 ry -13.97 rz 90 deg; joints [6.757, -81.654, 138.224, -171.92, 56.832, 161.591]
  MoveL 482 to (-31.75, -40.82, 11.93) mm, rotated rx 90 ry -15.85 rz 90 deg; joints [7.392, -81.409, 138.094, -171.175, 56.998, 159.322]
  MoveL 483 to (-30.82, -40.72, 11.58) mm, rotated rx 90 ry -17.72 rz 90 deg; joints [8.021, -81.133, 137.965, -170.444, 57.197, 157.068]
  MoveL 484 to (-29.89, -40.6, 11.23) mm, rotated rx 90 ry -19.6 rz 90 deg; joints [8.642, -80.827, 137.835, -169.729, 57.429, 154.831]
  MoveL 485 to (-28.96, -40.47, 10.88) mm, rotated rx 90 ry -21.47 rz 90 deg; joints [9.257, -80.492, 137.705, -169.029, 57.693, 152.611]
  MoveL 486 to (-28.03, -40.33, 10.54) mm, rotated rx 90 ry -23.35 rz 90 deg; joints [9.862, -80.127, 137.575, -168.346, 57.986, 150.41]
  MoveL 487 to (-27.1, -40.18, 10.21) mm, rotated rx 90 ry -25.23 rz 90 deg; joints [10.458, -79.734, 137.444, -167.682, 58.31, 148.229]
  MoveL 488 to (-26.25, -39.96, 9.78) mm, rotated rx 90 ry -27.66 rz 90 deg; joints [11.221, -79.203, 137.3, -166.847, 58.776, 145.432]
  MoveL 489 to (-25.39, -39.73, 9.36) mm, rotated rx 90 ry -30.1 rz 90 deg; joints [11.966, -78.625, 137.155, -166.046, 59.289, 142.672]
  MoveL 490 to (-24.54, -39.48, 8.95) mm, rotated rx 90 ry -32.53 rz 90 deg; joints [12.692, -78.003, 137.008, -165.28, 59.843, 139.951]
  MoveL 491 to (-23.68, -39.22, 8.55) mm, rotated rx 90 ry -34.97 rz 90 deg; joints [13.398, -77.337, 136.86, -164.55, 60.437, 137.27]
  MoveL 492 to (-22.92, -38.88, 8.09) mm, rotated rx 90 ry -37.9 rz 90 deg; joints [14.224, -76.493, 136.699, -163.718, 61.207, 134.094]
  MoveL 493 to (-22.15, -38.51, 7.64) mm, rotated rx 90 ry -40.83 rz 90 deg; joints [15.017, -75.59, 136.535, -162.939, 62.026, 130.976]
  MoveL 494 to (-21.38, -38.12, 7.22) mm, rotated rx 90 ry -43.76 rz 90 deg; joints [15.777, -74.631, 136.367, -162.215, 62.89, 127.919]
  MoveL 495 to (-20.61, -37.72, 6.81) mm, rotated rx 90 ry -46.7 rz 90 deg; joints [16.5, -73.619, 136.196, -161.545, 63.794, 124.919]
  MoveL 496 to (-19.73, -37.01, 6.2) mm, rotated rx 90 ry -51.49 rz 90 deg; joints [17.609, -71.877, 135.933, -160.559, 65.354, 120.138]
  MoveL 497 to (-18.85, -36.24, 5.64) mm, rotated rx 90 ry -56.28 rz 90 deg; joints [18.614, -70.013, 135.656, -159.71, 66.993, 115.498]
  MoveL 498 to (-17.96, -35.44, 5.15) mm, rotated rx 90 ry -61.07 rz 90 deg; joints [19.512, -68.039, 135.363, -158.991, 68.692, 110.984]
  MoveL 499 to (-17.41, -34.71, 4.78) mm, rotated rx 90 ry -65.25 rz 90 deg; joints [20.21, -66.25, 135.11, -158.462, 70.218, 107.144]
  MoveL 500 to (-16.86, -33.95, 4.47) mm, rotated rx 90 ry -69.42 rz 90 deg; joints [20.822, -64.397, 134.844, -158.022, 71.77, 103.38]
  MoveL 501 to (-16.31, -33.18, 4.21) mm, rotated rx 90 ry -73.6 rz 90 deg; joints [21.348, -62.49, 134.563, -157.668, 73.34, 99.681]
  MoveL 502 to (-15.76, -32.38, 4) mm, rotated rx 90 ry -77.78 rz 90 deg; joints [21.786, -60.538, 134.267, -157.395, 74.92, 96.039]
  MoveL 503 to (-15.3, -31.53, 3.85) mm, rotated rx 90 ry -82.19 rz 90 deg; joints [22.155, -58.441, 133.949, -157.19, 76.598, 92.239]
  MoveL 504 to (-14.85, -30.66, 3.77) mm, rotated rx 90 ry -86.61 rz 90 deg; joints [22.426, -56.316, 133.615, -157.069, 78.273, 88.477]
  MoveL 505 to (-14.39, -29.8, 3.75) mm, rotated rx 0 ry -90 rz 180 deg; joints [22.564, -54.654, 133.339, -157.035, 79.561, 85.61]
  MoveL 506 to (-13.93, -28.93, 3.75) mm, rotated rx 0 ry -90 rz 180 deg; joints [22.555, -54.577, 133.3, -157.047, 79.596, 85.626]
  MoveL 507 to (-12.22, -25.42, 3.75) mm, rotated rx 0 ry -90 rz 180 deg; joints [22.522, -54.267, 133.149, -157.091, 79.74, 85.695]
  MoveL 508 to (-9.48, -21.07, 3.75) mm, rotated rx 0 ry -90 rz 180 deg; joints [22.47, -53.867, 132.917, -157.156, 79.89, 85.771]
  MoveL 509 to (-5.64, -17.69, 3.75) mm, rotated rx 0 ry -90 rz 180 deg; joints [22.397, -53.513, 132.613, -157.233, 79.931, 85.804]
  MoveL 510 to (-1.07, -15.06, 3.75) mm, rotated rx 0 ry -90 rz 180 deg; joints [22.311, -53.196, 132.263, -157.318, 79.894, 85.806]
  MoveL 511 to (3.61, -12.69, 3.75) mm, rotated rx 0 ry -90 rz 180 deg; joints [22.223, -52.896, 131.905, -157.403, 79.834, 85.799]
  MoveL 512 to (8.27, -10.41, 3.75) mm, rotated rx 0 ry -90 rz 180 deg; joints [22.136, -52.606, 131.55, -157.486, 79.768, 85.789]
  MoveL 513 to (17.27, -5.84, 3.75) mm, rotated rx 0 ry -90 rz 180 deg; joints [21.971, -52.033, 130.858, -157.646, 79.646, 85.773]
  MoveL 514 to (25.94, -0.5, 3.75) mm, rotated rx 0 ry -90 rz 180 deg; joints [21.814, -51.415, 130.177, -157.801, 79.576, 85.777]
  MoveL 515 to (74.06, -0.5, 3.75) mm, rotated rx 0 ry -90 rz 180 deg; joints [20.979, -50.108, 126.654, -158.483, 77.452, 85.104]
  MoveL 516 to (82.73, -5.84, 3.75) mm, rotated rx 0 ry -90 rz 180 deg; joints [20.835, -50.23, 126.062, -158.57, 76.776, 84.869]
  MoveL 517 to (91.73, -10.41, 3.75) mm, rotated rx 0 ry -90 rz 180 deg; joints [20.687, -50.279, 125.432, -158.662, 76.13, 84.65]
  MoveL 518 to (96.39, -12.69, 3.75) mm, rotated rx 0 ry -90 rz 180 deg; joints [20.612, -50.295, 125.103, -158.708, 75.802, 84.54]
  MoveL 519 to (101.07, -15.06, 3.75) mm, rotated rx 0 ry -90 rz 180 deg; joints [20.536, -50.315, 124.772, -158.753, 75.468, 84.427]
  MoveL 520 to (105.64, -17.69, 3.75) mm, rotated rx 0 ry -90 rz 180 deg; joints [20.463, -50.353, 124.45, -158.794, 75.125, 84.312]
  MoveL 521 to (109.48, -21.07, 3.75) mm, rotated rx 0 ry -90 rz 180 deg; joints [20.402, -50.46, 124.187, -158.821, 74.774, 84.19]
  MoveL 522 to (112.22, -25.42, 3.75) mm, rotated rx 0 ry -90 rz 180 deg; joints [20.359, -50.662, 124.014, -158.828, 74.419, 84.061]
  MoveL 523 to (113.93, -28.93, 3.75) mm, rotated rx 0 ry -90 rz 180 deg; joints [20.332, -50.84, 123.911, -158.827, 74.154, 83.963]
  MoveL 524 to (114.39, -29.8, 3.75) mm, rotated rx 0 ry -90 rz 180 deg; joints [20.324, -50.883, 123.882, -158.827, 74.087, 83.938]
  MoveL 525 to (114.85, -30.66, 3.77) mm, rotated rx 90 ry -86.61 rz 90 deg; joints [20.182, -52.313, 124.073, -158.842, 72.916, 86.904]
  MoveL 526 to (115.3, -31.53, 3.85) mm, rotated rx 90 ry -82.19 rz 90 deg; joints [19.919, -54.143, 124.32, -158.933, 71.408, 90.804]
  MoveL 527 to (115.76, -32.38, 4) mm, rotated rx 90 ry -77.78 rz 90 deg; joints [19.566, -55.942, 124.554, -159.108, 69.902, 94.749]
  MoveL 528 to (116.31, -33.18, 4.21) mm, rotated rx 90 ry -73.6 rz 90 deg; joints [19.147, -57.602, 124.755, -159.355, 68.482, 98.53]
  MoveL 529 to (116.86, -33.95, 4.47) mm, rotated rx 90 ry -69.42 rz 90 deg; joints [18.65, -59.218, 124.944, -159.683, 67.076, 102.369]
  MoveL 530 to (117.42, -34.71, 4.78) mm, rotated rx 90 ry -65.25 rz 90 deg; joints [18.076, -60.781, 125.122, -160.096, 65.692, 106.275]
  MoveL 531 to (117.97, -35.44, 5.15) mm, rotated rx 90 ry -61.07 rz 90 deg; joints [17.425, -62.282, 125.289, -160.596, 64.338, 110.256]
  MoveL 532 to (118.85, -36.24, 5.64) mm, rotated rx 90 ry -56.28 rz 90 deg; joints [16.586, -63.909, 125.448, -161.284, 62.823, 114.924]
  MoveL 533 to (119.73, -37.01, 6.2) mm, rotated rx 90 ry -51.49 rz 90 deg; joints [15.654, -65.433, 125.593, -162.097, 61.372, 119.713]
  MoveL 534 to (120.61, -37.72, 6.81) mm, rotated rx 90 ry -46.7 rz 90 deg; joints [14.635, -66.843, 125.728, -163.038, 60, 124.631]
  MoveL 535 to (121.38, -38.12, 7.22) mm, rotated rx 90 ry -43.76 rz 90 deg; joints [13.967, -67.636, 125.787, -163.68, 59.198, 127.708]
  MoveL 536 to (122.15, -38.51, 7.64) mm, rotated rx 90 ry -40.83 rz 90 deg; joints [13.27, -68.379, 125.843, -164.371, 58.435, 130.837]
  MoveL 537 to (122.92, -38.88, 8.09) mm, rotated rx 90 ry -37.9 rz 90 deg; joints [12.546, -69.071, 125.896, -165.111, 57.715, 134.02]
  MoveL 538 to (123.68, -39.22, 8.55) mm, rotated rx 90 ry -34.97 rz 90 deg; joints [11.795, -69.711, 125.946, -165.899, 57.041, 137.253]
  MoveL 539 to (124.54, -39.48, 8.95) mm, rotated rx 90 ry -32.53 rz 90 deg; joints [11.152, -70.189, 125.969, -166.59, 56.513, 139.976]
  MoveL 540 to (125.39, -39.73, 9.36) mm, rotated rx 90 ry -30.1 rz 90 deg; joints [10.494, -70.628, 125.991, -167.312, 56.023, 142.733]
  MoveL 541 to (126.25, -39.96, 9.78) mm, rotated rx 90 ry -27.66 rz 90 deg; joints [9.822, -71.027, 126.011, -168.064, 55.571, 145.523]
  MoveL 542 to (127.1, -40.18, 10.21) mm, rotated rx 90 ry -25.23 rz 90 deg; joints [9.137, -71.385, 126.03, -168.844, 55.159, 148.345]
  MoveL 543 to (128.03, -40.33, 10.54) mm, rotated rx 90 ry -23.35 rz 90 deg; joints [8.6, -71.619, 126.023, -169.465, 54.864, 150.541]
  MoveL 544 to (128.96, -40.47, 10.88) mm, rotated rx 90 ry -21.47 rz 90 deg; joints [8.056, -71.827, 126.016, -170.099, 54.595, 152.752]
  MoveL 545 to (129.89, -40.6, 11.23) mm, rotated rx 90 ry -19.6 rz 90 deg; joints [7.507, -72.011, 126.007, -170.748, 54.353, 154.98]
  MoveL 546 to (130.82, -40.72, 11.58) mm, rotated rx 90 ry -17.72 rz 90 deg; joints [6.954, -72.168, 125.998, -171.408, 54.138, 157.221]
  MoveL 547 to (131.75, -40.82, 11.93) mm, rotated rx 90 ry -15.85 rz 90 deg; joints [6.397, -72.299, 125.989, -172.08, 53.951, 159.475]
  MoveL 548 to (132.68, -40.92, 12.28) mm, rotated rx 90 ry -13.97 rz 90 deg; joints [5.836, -72.405, 125.979, -172.761, 53.793, 161.741]
  MoveL 549 to (133.66, -40.97, 12.48) mm, rotated rx 90 ry -12.93 rz 90 deg; joints [5.523, -72.427, 125.937, -173.142, 53.707, 162.998]
  MoveL 550 to (134.64, -41.01, 12.68) mm, rotated rx 90 ry -11.89 rz 90 deg; joints [5.208, -72.441, 125.896, -173.527, 53.63, 164.26]
  MoveL 551 to (135.62, -41.05, 12.88) mm, rotated rx 90 ry -10.85 rz 90 deg; joints [4.894, -72.447, 125.854, -173.912, 53.562, 165.522]
  MoveL 552 to (136.6, -41.09, 13.08) mm, rotated rx 90 ry -9.81 rz 90 deg; joints [4.58, -72.444, 125.811, -174.3, 53.503, 166.788]
  MoveL 553 to (137.58, -41.12, 13.28) mm, rotated rx 90 ry -8.78 rz 90 deg; joints [4.265, -72.434, 125.769, -174.688, 53.453, 168.055]
  MoveL 554 to (138.56, -41.15, 13.48) mm, rotated rx 90 ry -7.74 rz 90 deg; joints [3.951, -72.415, 125.726, -175.077, 53.412, 169.323]
  MoveL 555 to (139.54, -41.15, 13.49) mm, rotated rx 90 ry -7.7 rz 90 deg; joints [3.936, -72.363, 125.651, -175.094, 53.389, 169.371]
  MoveL 556 to (140.52, -41.15, 13.5) mm, rotated rx 90 ry -7.66 rz 90 deg; joints [3.922, -72.311, 125.577, -175.111, 53.366, 169.417]
  MoveL 557 to (141.5, -41.15, 13.51) mm, rotated rx 90 ry -7.62 rz 90 deg; joints [3.907, -72.259, 125.502, -175.128, 53.342, 169.464]
  MoveL 558 to (142.49, -41.15, 13.52) mm, rotated rx 90 ry -7.59 rz 90 deg; joints [3.893, -72.206, 125.427, -175.144, 53.319, 169.51]
  MoveL 559 to (143.45, -41.12, 13.32) mm, rotated rx 90 ry -8.6 rz 90 deg; joints [4.191, -72.122, 125.32, -174.771, 53.313, 168.276]
  MoveL 560 to (144.41, -41.09, 13.12) mm, rotated rx 90 ry -9.61 rz 90 deg; joints [4.489, -72.03, 125.214, -174.4, 53.315, 167.041]
  MoveL 561 to (145.37, -41.06, 12.93) mm, rotated rx 90 ry -10.62 rz 90 deg; joints [4.785, -71.931, 125.107, -174.03, 53.325, 165.81]
  MoveL 562 to (146.33, -41.02, 12.73) mm, rotated rx 90 ry -11.63 rz 90 deg; joints [5.081, -71.824, 125, -173.662, 53.344, 164.579]
  MoveL 563 to (147.25, -40.93, 12.33) mm, rotated rx 90 ry -13.73 rz 90 deg; joints [5.696, -71.637, 124.86, -172.901, 53.434, 162.028]
  MoveL 564 to (148.16, -40.82, 11.93) mm, rotated rx 90 ry -15.83 rz 90 deg; joints [6.308, -71.418, 124.72, -172.151, 53.56, 159.487]
  MoveL 565 to (149.08, -40.7, 11.54) mm, rotated rx 90 ry -17.93 rz 90 deg; joints [6.913, -71.167, 124.579, -171.414, 53.72, 156.959]
  MoveL 566 to (150, -40.57, 11.14) mm, rotated rx 90 ry -20.04 rz 90 deg; joints [7.511, -70.886, 124.437, -170.691, 53.914, 154.448]
  MoveL 567 to (150, -40.2, 10.26) mm, rotated rx 90 ry -24.92 rz 90 deg; joints [8.884, -70.228, 124.271, -169.07, 54.54, 148.688]
  MoveL 568 to (150, -39.76, 9.41) mm, rotated rx 90 ry -29.8 rz 90 deg; joints [10.209, -69.409, 124.1, -167.555, 55.331, 143.043]
  MoveL 569 to (150, -39.25, 8.6) mm, rotated rx 90 ry -34.69 rz 90 deg; joints [11.477, -68.437, 123.924, -166.157, 56.271, 137.524]
  MoveL 570 to (150, -38.67, 7.83) mm, rotated rx 90 ry -39.57 rz 90 deg; joints [12.679, -67.319, 123.74, -164.889, 57.343, 132.143]
  MoveL 571 to (150, -38.03, 7.12) mm, rotated rx 90 ry -44.45 rz 90 deg; joints [13.805, -66.065, 123.549, -163.754, 58.533, 126.902]
  MoveL 572 to (150, -37.33, 6.47) mm, rotated rx 90 ry -49.33 rz 90 deg; joints [14.85, -64.683, 123.347, -162.754, 59.822, 121.799]
  MoveL 573 to (150, -36.58, 5.87) mm, rotated rx 90 ry -54.21 rz 90 deg; joints [15.808, -63.185, 123.135, -161.888, 61.196, 116.83]
  MoveL 574 to (150, -35.78, 5.35) mm, rotated rx 90 ry -59.1 rz 90 deg; joints [16.673, -61.582, 122.91, -161.153, 62.638, 111.987]
  MoveL 575 to (150, -34.94, 4.89) mm, rotated rx 90 ry -63.98 rz 90 deg; joints [17.44, -59.884, 122.671, -160.544, 64.134, 107.261]
  MoveL 576 to (150, -34.06, 4.51) mm, rotated rx 90 ry -68.86 rz 90 deg; joints [18.107, -58.104, 122.418, -160.057, 65.671, 102.638]
  MoveL 577 to (150, -33.15, 4.2) mm, rotated rx 90 ry -73.74 rz 90 deg; joints [18.671, -56.255, 122.15, -159.686, 67.238, 98.106]
  MoveL 578 to (150, -32.22, 3.97) mm, rotated rx 90 ry -78.62 rz 90 deg; joints [19.129, -54.348, 121.868, -159.425, 68.823, 93.652]
  MoveL 579 to (150, -31.27, 3.82) mm, rotated rx 90 ry -83.51 rz 90 deg; joints [19.48, -52.397, 121.57, -159.271, 70.415, 89.263]
  MoveL 580 to (150, -30.32, 3.75) mm, rotated rx 90 ry -88.39 rz 90 deg; joints [19.723, -50.415, 121.259, -159.218, 72.007, 84.925]
  MoveL 581 to (150, -29.36, 3.75) mm, rotated rx 0 ry -90 rz 180 deg; joints [19.779, -49.716, 121.149, -159.226, 72.565, 83.515]
  MoveL 582 to (150, -28.4, 3.75) mm, rotated rx 0 ry -90 rz 180 deg; joints [19.779, -49.655, 121.142, -159.232, 72.615, 83.536]
  MoveL 583 to (146.28, -29.22, 3.75) mm, rotated rx 0 ry -90 rz 180 deg; joints [19.834, -49.828, 121.436, -159.187, 72.734, 83.563]
  MoveL 584 to (142.22, -28.97, 3.75) mm, rotated rx 0 ry -90 rz 180 deg; joints [19.895, -49.943, 121.747, -159.145, 72.925, 83.617]
  MoveL 585 to (138.31, -27.66, 3.75) mm, rotated rx 0 ry -90 rz 180 deg; joints [19.955, -49.986, 122.039, -159.111, 73.164, 83.692]
  MoveL 586 to (135.78, -26.02, 3.75) mm, rotated rx 0 ry -90 rz 180 deg; joints [19.993, -49.961, 122.221, -159.093, 73.362, 83.758]
  MoveL 587 to (133.82, -23.81, 3.75) mm, rotated rx 0 ry -90 rz 180 deg; joints [20.023, -49.88, 122.355, -159.085, 73.565, 83.829]
  MoveL 588 to (132.64, -21.07, 3.75) mm, rotated rx 0 ry -90 rz 180 deg; joints [20.041, -49.74, 122.424, -159.088, 73.762, 83.901]
  MoveL 589 to (132.34, -17.66, 3.75) mm, rotated rx 0 ry -90 rz 180 deg; joints [20.046, -49.529, 122.419, -159.105, 73.956, 83.977]
  MoveL 590 to (133.11, -14.37, 3.75) mm, rotated rx 0 ry -90 rz 180 deg; joints [20.034, -49.291, 122.332, -159.132, 74.095, 84.036]
  MoveL 591 to (134.92, -11.65, 3.75) mm, rotated rx 0 ry -90 rz 180 deg; joints [20.006, -49.058, 122.17, -159.168, 74.158, 84.07]
  MoveL 592 to (137.54, -9.53, 3.75) mm, rotated rx 0 ry -90 rz 180 deg; joints [19.966, -48.84, 121.95, -159.209, 74.153, 84.081]
  MoveL 593 to (141.76, -7.46, 3.75) mm, rotated rx 0 ry -90 rz 180 deg; joints [19.902, -48.575, 121.607, -159.267, 74.073, 84.07]
  MoveL 594 to (146.15, -6.05, 3.75) mm, rotated rx 0 ry -90 rz 180 deg; joints [19.836, -48.349, 121.256, -159.323, 73.95, 84.043]
  MoveL 595 to (150, -5.07, 3.75) mm, rotated rx 0 ry -90 rz 180 deg; joints [19.779, -48.166, 120.949, -159.37, 73.827, 84.014]
  MoveL 596 to (134.08, 0, 3.75) mm, rotated rx 0 ry -90 rz 180 deg; joints [20.019, -48.326, 122.126, -159.223, 74.803, 84.32]
  MoveL 597 to (133.99, -2.31, 3.75) mm, rotated rx 0 ry -90 rz 180 deg; joints [20.021, -48.479, 122.155, -159.209, 74.688, 84.274]
  MoveL 598 to (133.12, -4.45, 3.75) mm, rotated rx 0 ry -90 rz 180 deg; joints [20.034, -48.645, 122.242, -159.188, 74.615, 84.242]
  MoveL 599 to (131.64, -6.32, 3.75) mm, rotated rx 0 ry -90 rz 180 deg; joints [20.057, -48.812, 122.373, -159.161, 74.584, 84.222]
  MoveL 600 to (128.64, -8.39, 3.75) mm, rotated rx 0 ry -90 rz 180 deg; joints [20.103, -49.039, 122.621, -159.115, 74.608, 84.217]
  MoveL 601 to (125.24, -9.27, 3.75) mm, rotated rx 0 ry -90 rz 180 deg; joints [20.155, -49.201, 122.889, -159.071, 74.713, 84.242]
  MoveL 602 to (120.92, -8.94, 3.75) mm, rotated rx 0 ry -90 rz 180 deg; joints [20.222, -49.31, 123.215, -159.023, 74.922, 84.304]
  MoveL 603 to (116.63, -8.26, 3.75) mm, rotated rx 0 ry -90 rz 180 deg; joints [20.289, -49.395, 123.535, -158.977, 75.148, 84.374]
  MoveL 604 to (112.36, -7.56, 3.75) mm, rotated rx 0 ry -90 rz 180 deg; joints [20.357, -49.476, 123.852, -158.93, 75.374, 84.444]
  MoveL 605 to (102.41, -5.59, 3.75) mm, rotated rx 0 ry -90 rz 180 deg; joints [20.515, -49.64, 124.585, -158.82, 75.92, 84.615]
  MoveL 606 to (93.68, -3.23, 3.75) mm, rotated rx 0 ry -90 rz 180 deg; joints [20.655, -49.736, 125.218, -158.723, 76.434, 84.781]
  MoveL 607 to (85.1, 0, 3.75) mm, rotated rx 0 ry -90 rz 180 deg; joints [20.796, -49.762, 125.828, -158.63, 76.99, 84.966]
  MoveL 608 to (14.9, 0, 3.75) mm, rotated rx 0 ry -90 rz 180 deg; joints [22.014, -51.666, 130.968, -157.634, 80.091, 85.95]
  MoveL 609 to (6.32, -3.23, 3.75) mm, rotated rx 0 ry -90 rz 180 deg; joints [22.173, -52.125, 131.618, -157.487, 80.277, 85.996]
  MoveL 610 to (-2.41, -5.59, 3.75) mm, rotated rx 0 ry -90 rz 180 deg; joints [22.336, -52.525, 132.266, -157.338, 80.519, 86.065]
  MoveL 611 to (-12.36, -7.56, 3.75) mm, rotated rx 0 ry -90 rz 180 deg; joints [22.525, -52.925, 132.994, -157.167, 80.833, 86.163]
  MoveL 612 to (-16.62, -8.26, 3.75) mm, rotated rx 0 ry -90 rz 180 deg; joints [22.607, -53.087, 133.304, -157.094, 80.975, 86.208]
  MoveL 613 to (-20.92, -8.94, 3.75) mm, rotated rx 0 ry -90 rz 180 deg; joints [22.69, -53.246, 133.615, -157.019, 81.12, 86.255]
  MoveL 614 to (-25.24, -9.27, 3.75) mm, rotated rx 0 ry -90 rz 180 deg; joints [22.774, -53.38, 133.923, -156.945, 81.286, 86.311]
  MoveL 615 to (-28.64, -8.39, 3.75) mm, rotated rx 0 ry -90 rz 180 deg; joints [22.841, -53.397, 134.154, -156.89, 81.488, 86.386]
  MoveL 616 to (-31.64, -6.32, 3.75) mm, rotated rx 0 ry -90 rz 180 deg; joints [22.9, -53.311, 134.344, -156.847, 81.745, 86.486]
  MoveL 617 to (-33.12, -4.45, 3.75) mm, rotated rx 0 ry -90 rz 180 deg; joints [22.929, -53.203, 134.428, -156.828, 81.924, 86.559]
  MoveL 618 to (-33.99, -2.31, 3.75) mm, rotated rx 0 ry -90 rz 180 deg; joints [22.946, -53.058, 134.467, -156.821, 82.093, 86.629]
  MoveL 619 to (-34.08, 0, 3.75) mm, rotated rx 0 ry -90 rz 180 deg; joints [22.948, -52.881, 134.448, -156.828, 82.238, 86.691]
  MoveL 620 to (-50, -5.07, 3.75) mm, rotated rx 0 ry -90 rz 180 deg; joints [23.268, -53.655, 135.616, -156.526, 82.618, 86.806]
  MoveL 621 to (-46.15, -6.05, 3.75) mm, rotated rx 0 ry -90 rz 180 deg; joints [23.19, -53.641, 135.358, -156.592, 82.39, 86.719]
  MoveL 622 to (-41.76, -7.46, 3.75) mm, rotated rx 0 ry -90 rz 180 deg; joints [23.101, -53.645, 135.065, -156.665, 82.113, 86.612]
  MoveL 623 to (-37.54, -9.53, 3.75) mm, rotated rx 0 ry -90 rz 180 deg; joints [23.017, -53.704, 134.791, -156.732, 81.802, 86.491]
  MoveL 624 to (-34.92, -11.65, 3.75) mm, rotated rx 0 ry -90 rz 180 deg; joints [22.965, -53.804, 134.629, -156.769, 81.558, 86.394]
  MoveL 625 to (-33.11, -14.37, 3.75) mm, rotated rx 0 ry -90 rz 180 deg; joints [22.929, -53.969, 134.528, -156.79, 81.311, 86.293]
  MoveL 626 to (-32.34, -17.66, 3.75) mm, rotated rx 0 ry -90 rz 180 deg; joints [22.913, -54.202, 134.504, -156.789, 81.074, 86.193]
  MoveL 627 to (-32.64, -21.07, 3.75) mm, rotated rx 0 ry -90 rz 180 deg; joints [22.919, -54.473, 134.557, -156.77, 80.874, 86.105]
  MoveL 628 to (-33.82, -23.81, 3.75) mm, rotated rx 0 ry -90 rz 180 deg; joints [22.943, -54.714, 134.664, -156.737, 80.752, 86.048]
  MoveL 629 to (-35.77, -26.02, 3.75) mm, rotated rx 0 ry -90 rz 180 deg; joints [22.982, -54.935, 134.82, -156.694, 80.696, 86.016]
  MoveL 630 to (-38.31, -27.66, 3.75) mm, rotated rx 0 ry -90 rz 180 deg; joints [23.032, -55.128, 135.012, -156.643, 80.698, 86.007]
  MoveL 631 to (-42.22, -28.97, 3.75) mm, rotated rx 0 ry -90 rz 180 deg; joints [23.11, -55.33, 135.298, -156.569, 80.78, 86.028]
  MoveL 632 to (-46.28, -29.22, 3.75) mm, rotated rx 0 ry -90 rz 180 deg; joints [23.192, -55.456, 135.584, -156.497, 80.933, 86.08]
  MoveL 633 to (-50, -28.4, 3.75) mm, rotated rx 0 ry -90 rz 180 deg; joints [23.268, -55.488, 135.838, -156.434, 81.142, 86.157]
  MoveL 634 to (-50, -28.4, -41.25) mm, rotated rx 0 ry -90 rz 180 deg; joints [25.363, -54.962, 134.423, -154.257, 80.487, 85.444]
  Sollgeschwindigkeit (200.0 mm/s)
  MoveL 635 to (-46.19, -34.34, -41.08) mm, rotated rx 90 ry -85.57 rz 90 deg; joints [25.074, -57.414, 134.524, -154.36, 78.343, 88.89]
  MoveL 636 to (-42.38, -43.28, -39.66) mm, rotated rx 90 ry -76.34 rz 90 deg; joints [24.205, -62.263, 134.925, -154.784, 74.229, 96.366]
  MoveL 637 to (-38.58, -51.88, -36.82) mm, rotated rx 90 ry -67.11 rz 90 deg; joints [22.861, -66.862, 135.233, -155.603, 70.145, 104.135]
  MoveL 638 to (-34.77, -59.91, -32.64) mm, rotated rx 90 ry -57.88 rz 90 deg; joints [21.056, -71.098, 135.452, -156.874, 66.177, 112.336]
  MoveL 639 to (-30.96, -67.17, -27.22) mm, rotated rx 90 ry -48.65 rz 90 deg; joints [18.81, -74.863, 135.598, -158.672, 62.436, 121.113]
  MoveL 640 to (-27.15, -73.46, -20.71) mm, rotated rx 90 ry -39.41 rz 90 deg; joints [16.156, -78.055, 135.69, -161.069, 59.058, 130.585]
  MoveL 641 to (-23.34, -78.62, -13.28) mm, rotated rx 90 ry -30.18 rz 90 deg; joints [13.148, -80.585, 135.752, -164.115, 56.206, 140.824]
  MoveL 642 to (-19.53, -82.53, -5.11) mm, rotated rx 90 ry -20.95 rz 90 deg; joints [9.857, -82.377, 135.805, -167.792, 54.054, 151.811]
  MoveL 643 to (-15.73, -85.08, 3.57) mm, rotated rx 90 ry -11.72 rz 90 deg; joints [6.377, -83.372, 135.864, -171.981, 52.764, 163.408]
  MoveL 644 to (-11.92, -86.2, 12.56) mm, rotated rx 90 ry -2.49 rz 90 deg; joints [2.818, -83.532, 135.934, -176.444, 52.455, 175.344]
  MoveL 645 to (-8.11, -86.25, 17.25) mm, rotated rx 90 ry 0 rz 90 deg; joints [1.735, -83.265, 135.762, -177.813, 52.518, 178.669]
  MoveL 646 to (-4.3, -86.25, 20.32) mm, rotated rx 90 ry 0 rz 90 deg; joints [1.564, -83.037, 135.497, -178.028, 52.476, 178.799]
  MoveL 647 to (-0.49, -86.25, 23.4) mm, rotated rx 90 ry 0 rz 90 deg; joints [1.394, -82.81, 135.231, -178.241, 52.434, 178.928]
  MoveL 648 to (3.32, -86.25, 26.48) mm, rotated rx 90 ry 0 rz 90 deg; joints [1.225, -82.582, 134.964, -178.454, 52.391, 179.056]
  MoveL 649 to (7.12, -86.25, 29.56) mm, rotated rx 90 ry 0 rz 90 deg; joints [1.057, -82.355, 134.695, -178.665, 52.348, 179.184]
  MoveL 650 to (10.93, -86.25, 32.63) mm, rotated rx 90 ry 0 rz 90 deg; joints [0.891, -82.128, 134.425, -178.874, 52.303, 179.312]
  MoveL 651 to (14.74, -86.25, 35.71) mm, rotated rx 90 ry 0 rz 90 deg; joints [0.725, -81.9, 134.155, -179.083, 52.258, 179.439]
  MoveL 652 to (18.55, -86.25, 38.79) mm, rotated rx 90 ry 0 rz 90 deg; joints [0.561, -81.673, 133.883, -179.29, 52.212, 179.565]
  MoveL 653 to (22.36, -86.25, 41.87) mm, rotated rx 90 ry 0 rz 90 deg; joints [0.398, -81.446, 133.609, -179.496, 52.165, 179.691]
  MoveL 654 to (26.16, -86.25, 44.94) mm, rotated rx 90 ry 0 rz 90 deg; joints [0.236, -81.219, 133.335, -179.701, 52.117, 179.816]
  MoveL 655 to (29.97, -85.55, 53.86) mm, rotated rx 90 ry 9.06 rz 90 deg; joints [-3.069, -80.254, 133.26, 176.159, 53.068, -168.631]
  MoveL 656 to (33.78, -83.41, 62.65) mm, rotated rx 90 ry 18.29 rz 90 deg; joints [-6.25, -78.503, 133.169, 172.353, 54.907, -157.296]
  MoveL 657 to (37.59, -79.89, 70.99) mm, rotated rx 90 ry 27.52 rz 90 deg; joints [-9.152, -76.021, 133.029, 169.127, 57.481, -146.582]
  MoveL 658 to (41.4, -75.07, 78.66) mm, rotated rx 90 ry 36.75 rz 90 deg; joints [-11.7, -72.878, 132.81, 166.543, 60.619, -136.551]
  Sollgeschwindigkeit (50.0 mm/s)
  MoveL 659 to (41.4, -39.01, 51.73) mm, rotated rx 90 ry 36.75 rz 90 deg; joints [-10.364, -70.867, 133.75, 168.389, 63.362, -137.983]
  MoveL 660 to (40.45, -39.05, 51.68) mm, rotated rx 90 ry 36.41 rz 90 deg; joints [-10.295, -71.022, 133.823, 168.458, 63.274, -138.339]
  MoveL 661 to (39.49, -39.09, 51.62) mm, rotated rx 90 ry 36.08 rz 90 deg; joints [-10.225, -71.177, 133.895, 168.528, 63.187, -138.694]
  MoveL 662 to (38.54, -39.13, 51.57) mm, rotated rx 90 ry 35.74 rz 90 deg; joints [-10.154, -71.331, 133.967, 168.598, 63.1, -139.051]
  MoveL 663 to (37.59, -39.17, 51.52) mm, rotated rx 90 ry 35.4 rz 90 deg; joints [-10.083, -71.485, 134.039, 168.67, 63.013, -139.408]
  MoveL 664 to (36.63, -39.21, 51.46) mm, rotated rx 90 ry 35.06 rz 90 deg; joints [-10.011, -71.638, 134.111, 168.742, 62.927, -139.764]
  MoveL 665 to (35.68, -39.25, 51.41) mm, rotated rx 90 ry 34.72 rz 90 deg; joints [-9.939, -71.791, 134.182, 168.815, 62.84, -140.122]
  MoveL 666 to (34.73, -39.28, 51.35) mm, rotated rx 90 ry 34.38 rz 90 deg; joints [-9.866, -71.943, 134.254, 168.888, 62.754, -140.481]
  MoveL 667 to (33.78, -39.32, 51.3) mm, rotated rx 90 ry 34.04 rz 90 deg; joints [-9.792, -72.095, 134.325, 168.963, 62.668, -140.84]
  MoveL 668 to (32.83, -39.36, 51.24) mm, rotated rx 90 ry 33.7 rz 90 deg; joints [-9.718, -72.247, 134.396, 169.038, 62.583, -141.2]
  MoveL 669 to (31.88, -39.44, 51.12) mm, rotated rx 90 ry 32.99 rz 90 deg; joints [-9.551, -72.511, 134.467, 169.207, 62.377, -141.96]
  MoveL 670 to (30.93, -39.51, 51.01) mm, rotated rx 90 ry 32.27 rz 90 deg; joints [-9.381, -72.773, 134.536, 169.379, 62.174, -142.722]
  MoveL 671 to (29.98, -39.59, 50.89) mm, rotated rx 90 ry 31.56 rz 90 deg; joints [-9.21, -73.032, 134.606, 169.554, 61.973, -143.488]
  MoveL 672 to (29.03, -39.66, 50.77) mm, rotated rx 90 ry 30.85 rz 90 deg; joints [-9.036, -73.288, 134.674, 169.732, 61.774, -144.256]
  MoveL 673 to (28.08, -39.73, 50.65) mm, rotated rx 90 ry 30.13 rz 90 deg; joints [-8.86, -73.54, 134.742, 169.914, 61.577, -145.027]
  MoveL 674 to (27.13, -39.8, 50.53) mm, rotated rx 90 ry 29.42 rz 90 deg; joints [-8.682, -73.79, 134.81, 170.099, 61.383, -145.801]
  MoveL 675 to (26.18, -39.87, 50.4) mm, rotated rx 90 ry 28.71 rz 90 deg; joints [-8.501, -74.036, 134.877, 170.287, 61.191, -146.579]
  MoveL 676 to (25.23, -39.93, 50.28) mm, rotated rx 90 ry 27.99 rz 90 deg; joints [-8.319, -74.279, 134.943, 170.479, 61.002, -147.36]
  MoveL 677 to (24.28, -40, 50.16) mm, rotated rx 90 ry 27.28 rz 90 deg; joints [-8.134, -74.519, 135.009, 170.674, 60.815, -148.143]
  MoveL 678 to (23.52, -40.11, 49.93) mm, rotated rx 90 ry 25.99 rz 90 deg; joints [-7.788, -74.894, 135.056, 171.04, 60.465, -149.566]
  MoveL 679 to (22.76, -40.22, 49.7) mm, rotated rx 90 ry 24.7 rz 90 deg; joints [-7.436, -75.258, 135.102, 171.416, 60.124, -151]
  MoveL 680 to (22, -40.32, 49.47) mm, rotated rx 90 ry 23.41 rz 90 deg; joints [-7.078, -75.61, 135.146, 171.803, 59.793, -152.445]
  MoveL 681 to (21.03, -40.58, 48.81) mm, rotated rx 90 ry 19.82 rz 90 deg; joints [-6.046, -76.461, 135.179, 172.936, 58.911, -156.516]
  MoveL 682 to (20.05, -40.8, 48.15) mm, rotated rx 90 ry 16.23 rz 90 deg; joints [-4.974, -77.213, 135.203, 174.14, 58.125, -160.663]
  MoveL 683 to (19.55, -40.98, 47.47) mm, rotated rx 90 ry 12.69 rz 90 deg; joints [-3.881, -77.827, 135.187, 175.394, 57.443, -164.823]
  MoveL 684 to (19.04, -41.11, 46.79) mm, rotated rx 90 ry 9.15 rz 90 deg; joints [-2.76, -78.339, 135.165, 176.704, 56.87, -169.042]
  MoveL 685 to (18.53, -41.2, 46.1) mm, rotated rx 90 ry 5.62 rz 90 deg; joints [-1.615, -78.744, 135.139, 178.061, 56.41, -173.312]
  MoveL 686 to (18.17, -41.25, 45.27) mm, rotated rx 90 ry 1.37 rz 90 deg; joints [-0.22, -79.074, 135.085, 179.734, 56.011, -178.479]
  MoveL 687 to (17.82, -41.25, 44.44) mm, rotated rx 90 ry 0 rz 90 deg; joints [0.264, -79.161, 135.084, -179.681, 55.924, 179.821]
  MoveL 688 to (17.47, -41.25, 43.6) mm, rotated rx 90 ry 0 rz 90 deg; joints [0.308, -79.181, 135.11, -179.628, 55.929, 179.791]
  MoveL 689 to (16.87, -41.25, 40.01) mm, rotated rx 90 ry 0 rz 90 deg; joints [0.497, -79.214, 135.152, -179.4, 55.939, 179.664]
  MoveL 690 to (17.29, -41.25, 36.56) mm, rotated rx 90 ry 0 rz 90 deg; joints [0.679, -79.188, 135.118, -179.181, 55.933, 179.541]
  MoveL 691 to (18.81, -41.25, 33.72) mm, rotated rx 90 ry 0 rz 90 deg; joints [0.827, -79.098, 135.004, -179.001, 55.91, 179.44]
  MoveL 692 to (21.87, -41.25, 30.71) mm, rotated rx 90 ry 0 rz 90 deg; joints [0.983, -78.921, 134.777, -178.813, 55.862, 179.334]
  MoveL 693 to (24.9, -41.25, 27.7) mm, rotated rx 90 ry 0 rz 90 deg; joints [1.137, -78.745, 134.551, -178.625, 55.814, 179.228]
  MoveL 694 to (27.3, -41.25, 24.26) mm, rotated rx 90 ry 0 rz 90 deg; joints [1.314, -78.603, 134.369, -178.411, 55.776, 179.106]
  MoveL 695 to (29.82, -41.25, 19.45) mm, rotated rx 90 ry 0 rz 90 deg; joints [1.561, -78.453, 134.175, -178.111, 55.737, 178.936]
  MoveL 696 to (30.23, -41.25, 18.61) mm, rotated rx 90 ry 0 rz 90 deg; joints [1.604, -78.429, 134.144, -178.059, 55.73, 178.907]
  MoveL 697 to (30.63, -41.25, 17.77) mm, rotated rx 90 ry 0 rz 90 deg; joints [1.647, -78.405, 134.112, -178.007, 55.724, 178.877]
  MoveL 698 to (31.03, -41.25, 16.94) mm, rotated rx 90 ry 0 rz 90 deg; joints [1.69, -78.38, 134.081, -177.955, 55.718, 178.848]
  MoveL 699 to (31.43, -41.25, 16.1) mm, rotated rx 90 ry 0 rz 90 deg; joints [1.733, -78.356, 134.05, -177.903, 55.712, 178.818]
  MoveL 700 to (31.84, -41.25, 15.26) mm, rotated rx 90 ry 0 rz 90 deg; joints [1.776, -78.332, 134.018, -177.851, 55.705, 178.789]
  MoveL 701 to (32.24, -41.23, 14.42) mm, rotated rx 90 ry -2.95 rz 90 deg; joints [2.756, -78.366, 133.893, -176.658, 55.572, 175.159]
  MoveL 702 to (32.68, -41.15, 13.54) mm, rotated rx 90 ry -7.48 rz 90 deg; joints [4.244, -78.286, 133.713, -174.851, 55.535, 169.601]
  MoveL 703 to (33.12, -41, 12.66) mm, rotated rx 90 ry -12.01 rz 90 deg; joints [5.722, -78.033, 133.531, -173.067, 55.694, 164.07]
  MoveL 704 to (33.56, -40.78, 11.8) mm, rotated rx 90 ry -16.54 rz 90 deg; joints [7.182, -77.61, 133.348, -171.331, 56.044, 158.593]
  MoveL 705 to (34, -40.5, 10.96) mm, rotated rx 90 ry -21.07 rz 90 deg; joints [8.611, -77.021, 133.163, -169.665, 56.575, 153.196]
  MoveL 706 to (34.44, -40.15, 10.14) mm, rotated rx 90 ry -25.6 rz 90 deg; joints [10.001, -76.271, 132.977, -168.087, 57.275, 147.896]
  MoveL 707 to (34.88, -39.73, 9.35) mm, rotated rx 90 ry -30.13 rz 90 deg; joints [11.341, -75.366, 132.787, -166.612, 58.133, 142.71]
  MoveL 708 to (35.31, -39.27, 8.63) mm, rotated rx 90 ry -34.51 rz 90 deg; joints [12.582, -74.35, 132.599, -165.293, 59.096, 137.811]
  MoveL 709 to (35.75, -38.76, 7.94) mm, rotated rx 90 ry -38.89 rz 90 deg; joints [13.762, -73.203, 132.405, -164.086, 60.178, 133.037]
  MoveL 710 to (36.18, -38.19, 7.29) mm, rotated rx 90 ry -43.28 rz 90 deg; joints [14.874, -71.932, 132.205, -162.994, 61.364, 128.385]
  MoveL 711 to (36.62, -37.58, 6.68) mm, rotated rx 90 ry -47.66 rz 90 deg; joints [15.914, -70.546, 131.998, -162.017, 62.64, 123.857]
  MoveL 712 to (37.01, -36.97, 6.17) mm, rotated rx 90 ry -51.71 rz 90 deg; joints [16.807, -69.169, 131.797, -161.215, 63.888, 119.773]
  MoveL 713 to (37.41, -36.33, 5.7) mm, rotated rx 90 ry -55.77 rz 90 deg; joints [17.63, -67.709, 131.588, -160.509, 65.192, 115.787]
  MoveL 714 to (37.8, -35.66, 5.28) mm, rotated rx 90 ry -59.82 rz 90 deg; joints [18.382, -66.173, 131.369, -159.894, 66.54, 111.888]
  MoveL 715 to (38.19, -34.95, 4.9) mm, rotated rx 90 ry -63.87 rz 90 deg; joints [19.059, -64.567, 131.139, -159.367, 67.926, 108.072]
  MoveL 716 to (38.52, -34.24, 4.58) mm, rotated rx 90 ry -67.84 rz 90 deg; joints [19.649, -62.942, 130.906, -158.935, 69.309, 104.413]
  MoveL 717 to (38.85, -33.51, 4.31) mm, rotated rx 90 ry -71.8 rz 90 deg; joints [20.164, -61.265, 130.663, -158.58, 70.712, 100.816]
  MoveL 718 to (39.18, -32.77, 4.1) mm, rotated rx 90 ry -75.76 rz 90 deg; joints [20.605, -59.546, 130.407, -158.299, 72.128, 97.274]
  MoveL 719 to (39.51, -32.01, 3.93) mm, rotated rx 90 ry -79.73 rz 90 deg; joints [20.969, -57.791, 130.14, -158.091, 73.552, 93.777]
  MoveL 720 to (39.83, -31.19, 3.81) mm, rotated rx 90 ry -83.92 rz 90 deg; joints [21.272, -55.904, 129.846, -157.946, 75.063, 90.116]
  MoveL 721 to (40.16, -30.37, 3.76) mm, rotated rx 90 ry -88.12 rz 90 deg; joints [21.489, -53.995, 129.541, -157.875, 76.57, 86.488]
  MoveL 722 to (40.48, -29.55, 3.75) mm, rotated rx 0 ry -90 rz 180 deg; joints [21.555, -53.097, 129.384, -157.873, 77.262, 84.877]
  MoveL 723 to (40.8, -28.72, 3.75) mm, rotated rx 0 ry -90 rz 180 deg; joints [21.549, -53.03, 129.354, -157.882, 77.297, 84.893]
  MoveL 724 to (42.19, -25.66, 3.75) mm, rotated rx 0 ry -90 rz 180 deg; joints [21.525, -52.773, 129.228, -157.918, 77.416, 84.949]
  MoveL 725 to (44.08, -22.58, 3.75) mm, rotated rx 0 ry -90 rz 180 deg; joints [21.492, -52.501, 129.064, -157.961, 77.514, 84.998]
  MoveL 726 to (46.71, -19.5, 3.75) mm, rotated rx 0 ry -90 rz 180 deg; joints [21.446, -52.208, 128.846, -158.014, 77.578, 85.036]
  MoveL 727 to (48.43, -18.08, 3.75) mm, rotated rx 0 ry -90 rz 180 deg; joints [21.416, -52.059, 128.708, -158.045, 77.586, 85.047]
  MoveL 728 to (50, -17.29, 3.75) mm, rotated rx 0 ry -90 rz 180 deg; joints [21.388, -51.959, 128.586, -158.071, 77.563, 85.045]
  MoveL 729 to (51.57, -18.08, 3.75) mm, rotated rx 0 ry -90 rz 180 deg; joints [21.361, -51.969, 128.478, -158.089, 77.451, 85.005]
  MoveL 730 to (53.29, -19.5, 3.75) mm, rotated rx 0 ry -90 rz 180 deg; joints [21.332, -52.021, 128.364, -158.106, 77.295, 84.949]
  MoveL 731 to (55.92, -22.58, 3.75) mm, rotated rx 0 ry -90 rz 180 deg; joints [21.286, -52.16, 128.196, -158.126, 77.006, 84.842]
  MoveL 732 to (57.81, -25.66, 3.75) mm, rotated rx 0 ry -90 rz 180 deg; joints [21.254, -52.32, 128.082, -158.135, 76.748, 84.744]
  MoveL 733 to (59.2, -28.72, 3.75) mm, rotated rx 0 ry -90 rz 180 deg; joints [21.23, -52.492, 128.003, -158.138, 76.514, 84.654]
  MoveL 734 to (59.52, -29.55, 3.75) mm, rotated rx 0 ry -90 rz 180 deg; joints [21.224, -52.54, 127.986, -158.137, 76.453, 84.631]
  MoveL 735 to (59.84, -30.37, 3.76) mm, rotated rx 90 ry -88.12 rz 90 deg; joints [21.148, -53.401, 128.094, -158.146, 75.746, 86.242]
  MoveL 736 to (60.17, -31.19, 3.81) mm, rotated rx 90 ry -83.92 rz 90 deg; joints [20.923, -55.251, 128.349, -158.219, 74.243, 89.885]
  MoveL 737 to (60.49, -32.01, 3.93) mm, rotated rx 90 ry -79.73 rz 90 deg; joints [20.614, -57.077, 128.593, -158.366, 72.738, 93.562]
  MoveL 738 to (60.82, -32.77, 4.1) mm, rotated rx 90 ry -75.76 rz 90 deg; joints [20.243, -58.77, 128.809, -158.577, 71.319, 97.074]
  MoveL 739 to (61.15, -33.51, 4.31) mm, rotated rx 90 ry -71.8 rz 90 deg; joints [19.798, -60.426, 129.014, -158.86, 69.91, 100.634]
  MoveL 740 to (61.48, -34.24, 4.58) mm, rotated rx 90 ry -67.84 rz 90 deg; joints [19.28, -62.037, 129.208, -159.216, 68.517, 104.25]
  MoveL 741 to (61.81, -34.95, 4.9) mm, rotated rx 90 ry -63.87 rz 90 deg; joints [18.69, -63.596, 129.39, -159.65, 67.145, 107.929]
